(* IEC 61131-3 sources: 2026_Projet_YGO_ExcavatriceDragage/CODE/J_SUPERVISION, 7 files *)

(* ---- GVL_Troubleshooting.st ---- *)
(* ═══════════════════════════════════════════════════════════════
   🕵️‍♂️ GVL_Troubleshooting — GVL Globale de Recherche de Pannes (Orientée Fonctions & Contexte)
   ───────────────────────────────────────────────────────────────
   ⚙️ Emplacement : CODE/J_SUPERVISION/GVL_Troubleshooting.st
   🎨 Structurée par CONTEXTE GLOBAL MACHINE + FONCTIONS MÉTIER (Utilisation Opérateur).
   💬 Permet de localiser en 3 secondes l'environnement et le blocage d'une action.
   ═══════════════════════════════════════════════════════════════ *)
{attribute 'qualified_only'}
VAR_GLOBAL
    A_ContexteMachineGlobal : ST_ChainContextGlobal; // 🌐 0. Contexte Global Machine (Mode, Simu, Commande, Bypass)
    B_Inputs                : ST_HardwareImage;     // 📥 1. Image complète des entrées réelles / qualifiées / simulées
    C_Safety                : ST_SafetyChecklist;   // 🛡️ 2. Diagnostic chronologique Chaîne de Sécurité & Réarmement AU
    D_Joystick              : ST_JoystickChecklist; // 🕹️ 3. Diagnostic chronologique Bus CANopen & Homme-Mort Joystick
    E_HomingM1              : ST_HomingChecklist;   // 🎯 4. Diagnostic chronologique Homing M1 (Treuil Retenue)
    F_HomingM2              : ST_HomingChecklist;   // 🎯 5. Diagnostic chronologique Homing M2 (Treuil Benne)
    G_CycleSemiAuto         : ST_ChainCycleSemiAuto;  // 🔄 6. Séquenceur de Cycle Semi-Automatique (X0 à X13)
    H_LevageSynchroniseM1M2 : ST_ChainWinchSync;     // 🛗 7. Levage Synchronisé M1+M2 (Mode Couplé Nominal)
    I_LevageUnitaireM1      : ST_ChainWinch;         // 🛗 8. Levage Unitaire M1 (Treuil Retenue)
    J_LevageUnitaireM2      : ST_ChainWinch;         // 🛗 9. Levage Unitaire M2 (Treuil Benne)
    K_BenneOuvertureFermeture: ST_ChainBucket;        // 🪣 10. Ouverture / Fermeture Benne
    L_TranslationPontM3     : ST_ChainTranslation;   // ↔️ 11. Translation Pont M3 (Variateur AC600)
    // M_Réserve
    N_MotionM1              : ST_MotionChecklist;   // ⚙️ 13. Diagnostic chronologique Mouvement M1 (Treuil Retenue)
    O_MotionM2              : ST_MotionChecklist;   // ⚙️ 14. Diagnostic chronologique Mouvement M2 (Treuil Benne)
    P_MotionM3              : ST_MotionChecklist;   // ⚙️ 15. Diagnostic chronologique Mouvement M3 (Translation)

    // 🕵️ Trace de blocage terrain (cause priorisée + horodatage) — produite par PRG_04/05
    Q_TraceWinchM1          : ST_TraceWinch;        // 🕵️ 16. Trace blocage treuil M1 (cause priorisée + horodatage)
    R_TraceWinchM2          : ST_TraceWinch;        // 🕵️ 17. Trace blocage treuil M2 (cause priorisée + horodatage)
    S_TraceTranslation      : ST_TraceTranslation;  // ↔️ 18. Trace blocage translation M3 (cause priorisée + horodatage)
    T_Permits : ST_PermitVisibilityHMI; // Vue unique IHM/terrain des permis canoniques
END_VAR

(* ---- FB_AntiFlickerText.st ---- *)
(* ═══════════════════════════════════════════════════════════════
   🧊 FB_AntiFlickerText — Lissage anti-clignotement d'un texte IHM
   ───────────────────────────────────────────────────────────────
   📄 Doc : DOC/AF/AF_Partie-07_Interface_IHM_v2.3.md §5.3
   🎯 Responsabilité : maintient un texte warning/état un temps minimum
      avant de laisser le contenu changer, et laisse passer en direct
      (sans maintien) les messages critiques (défauts AU/puissance).
   🛡️ Sécurité : l'action de sécurité reste instantanée — ce FB ne
      retarde jamais un texte, il ne fait que stabiliser l'affichage.
      Il n'a aucun effet sur la machine.
   ═══════════════════════════════════════════════════════════════ *)
FUNCTION_BLOCK PUBLIC FB_AntiFlickerText
VAR_INPUT
    NewText      : STRING(120);  (* --> [CMD] Texte candidat à afficher *)
    ForceInstant : BOOL;         (* --> [CMD] TRUE = afficher immédiatement (défaut critique), sans maintien *)
    HoldTime     : TIME := T#500ms; (* --> [CFG] Durée de maintien min avant changement (AF-07 §5.3) *)
END_VAR
VAR_OUTPUT
    Text         : STRING(120);  (* <-- [STAT] Texte stabilisé exposé à l'IHM *)
END_VAR
VAR
    TonHold      : TON;   (* . [LOC] Temporisation de maintien *)
END_VAR

{region "§1 Lissage anti-clignotement"}
// Défaut critique : affichage immédiat, le TON est remis à zéro (aucune latence).
IF ForceInstant THEN
    Text := NewText;
    TonHold(IN := FALSE);
ELSE
    // Warning / état : le texte ne change qu'après maintien min (HoldTime).
    // Un signal qui oscille plus vite que HoldTime → texte stable.
    TonHold(IN := (NewText <> Text), PT := HoldTime);
    IF TonHold.Q THEN
        Text := NewText;
    END_IF;
END_IF;
{endregion}

(* ---- FB_CfgT330Normalizer.st ---- *)
(* ═══════════════════════════════════════════════════════════════
   🔧 FB_CfgT330Normalizer — Normalisation des réglages HAUT (T330)
   ───────────────────────────────────────────────────────────────
   🎯 Rôle : ramener DANS SON DOMAINE le couple de réglages de fin de
             course HAUT — FDC logiciel (CfgCableLimitAscent_M) et cote
             TOP homing (CfgTopSensorPos_M) — plus le plancher du
             ralentissement haut (WinchSlowdownDistanceTop_M), puis
             signaler la correction à l'IHM.
   📄 Doc : DOC/WFLOW/AUDITS/DESIGN/PLAN_T330_C3_INVARIANT_HAUT_v1.0.md (plan C3 v1.3, §2/§4)
            DOC/WFLOW/AUDITS/DESIGN/CADRAGE_T330_INVARIANT_HAUT_v1.0.md
   🛡️ Sécurité : une valeur de réglage HORS DOMAINE resterait hors domaine
             indéfiniment sans ce bloc (contre-exemple Q21 bis : FDC=9,50 m +
             TOP=12,00 m, où Δ=2,50 m ≥ 1,00 m n'active AUCUNE règle Δ).
             ⇒ R0 (clamp absolu) est INCONDITIONNELLE et EN AMONT de la règle Δ.
             Ce FB ne commande AUCUN mouvement : il corrige de la configuration.
   🧩 Dépendances : ST_WinchCfg (CfgTopSensorPos_M) · ST_CommunCfg
             (CfgCableLimitAscent_M, WinchSlowdownDistanceTop_M).
   ⚠️ Ordre d'appel : AVANT les ponts de persistance (PRG_07_Supervision §2).
             Le pont écrit la valeur CORRIGÉE dans le MÊME scan (option A / Q23)
             ⇒ aucune fenêtre NVRAM. Les mémoires internes sont amorcées depuis
             ces valeurs RESTAURÉES, jamais depuis les défauts du DUT (piège P2).
   ═══════════════════════════════════════════════════════════════ *)

FUNCTION_BLOCK FB_CfgT330Normalizer
VAR_INPUT
    // === CONTRAT STANDARD (Enable) ===
    Enable              : BOOL;  // 🟢 Autorise la normalisation (ponts de config RESTAURÉS)

    // === CONTEXTE MACHINE ===
    InHoming            : BOOL;  // 🎯 Homing en cours : cycle machine COMPLET (HX0..HX6) OU transaction de preset, M1 ou M2
END_VAR

VAR_IN_OUT
    // === RÉGLAGES HAUT À NORMALISER (référence — jamais de copie) ===
    WinchCfgM1          : ST_WinchCfg;   // 🔧 M1 = MAÎTRE du capteur haut : porte CfgTopSensorPos_M
    CommunCfg           : ST_CommunCfg;  // 🔧 Commun M1/M2 : porte CfgCableLimitAscent_M + WinchSlowdownDistanceTop_M
END_VAR

VAR_OUTPUT
    // === CONTRAT STANDARD (Ready) ===
    Ready               : BOOL;  // 🟢 Normalisation armée ce scan (Enable ET mémoires amorcées)

    // === DIAGNOSTIC / IHM ===
    Corrected           : BOOL;  // 🔧 Une correction T330 a eu lieu CE scan (impulsion d'un seul scan)
    CorrectedHeld       : BOOL;  // 🔧 Maintien du message T330 (fenêtre IHM — 1 scan serait invisible)
END_VAR

VAR CONSTANT
    // === T330 (Q1/Q2) — RÈGLES D'INGÉNIERIE, PAS DES COTES MÉTIER ===
    // NON persistantes et NON IHM (AC3) : jamais exposées, jamais RETAIN.
    CST_T330ReserveMinMargin_M : REAL := 0.40;   // Réserve minimale FDC logiciel haut / TOP homing (decision humaine, ex-1.00m)
    CST_T330SlowdownTopMin_M   : REAL := 0.50;   // Plancher du ralentissement haut (Q1)
    CST_T330FdcMin_M           : REAL := 0.00;   // Borne basse FDC (Q21)
    CST_T330FdcMax_M           : REAL := 9.60;   // Borne haute FDC (Q21/C1 : TOP<=10 et Delta>=0.4 => FDC<=9.6)
    CST_T330TopMin_M           : REAL := 1.00;   // Borne basse TOP (Q21)
    CST_T330TopMax_M           : REAL := 10.00;  // Borne haute TOP (Q21)
END_VAR

VAR
    // === T330 — MÉMOIRES NON PERSISTANTES (AC3 : ni IHM, ni RETAIN) ===
    T330PrevInit               : BOOL;  // . [LOC] Seed des mémoires effectué depuis les valeurs RESTAURÉES
    T330PrevTopSensorPos_M     : REAL;  // . [LOC] Valeur précédente TOP (détection du champ modifié par l'opérateur)
    T330PrevCableLimitAscent_M : REAL;  // . [LOC] Valeur précédente FDC (détection du champ modifié par l'opérateur)
    T330MsgHold                : TOF;   // . [LOC] Maintien du message T330 (un scan de 10 ms serait invisible à l'IHM)
END_VAR

// ═══════════════════════════════════════════════════════════════════════════════
// 🔧 T330 — COHÉRENCE DES RÉGLAGES HAUT (Q1/Q2) · plan C3 v1.3
// ───────────────────────────────────────────────────────────────────────────────
// ORDRE IMPOSÉ (Q21 bis) :  (1) R0 clamp ABSOLU inconditionnel, FDC et TOP séparément
//                        puis (2) règle Delta >= 1,00 m / slowdown >= 0,50 m.
// OPTION A (Q23) : ce bloc s'exécute AVANT les ponts de persistance, qui écrivent la
//                  valeur CORRIGÉE dans le MÊME scan (aucune fenêtre NVRAM). La
//                  référence est donc lue sur GVL_IHM.Cfg — l'état que les ponts
//                  tiennent à jour, et NON directement la NVRAM.
// AC3 : AUCUNE variable persistante ni IHM nouvelle — constantes CST_* et mémoires
//       locales uniquement. Jamais de champ de fin de course supplémentaire.
// C2/Q22 : R2 (correction du TOP) est INHIBÉE pendant le homing — sur le CYCLE COMPLET
//          (HX0..HX6), pas seulement la transaction de preset (~50 ms). Aucune mémoire
//          d'intention : au retour, si la config est toujours invalide, le REPLI NIVEAU
//          ci-dessous applique Q17 (préserver le TOP, corriger le FDC).
// ═══════════════════════════════════════════════════════════════════════════════
{region "🔧 T330 NORMALISATION"}
Corrected := FALSE;
Ready := FALSE;

// Inhibée tant que les ponts n'ont pas RESTAURÉ (sinon les défauts DUT seraient pris
// pour une saisie opérateur — piège P2 du cadrage).
IF Enable THEN

    // Seed des mémoires depuis les valeurs RESTAURÉES (jamais depuis les défauts DUT).
    IF NOT T330PrevInit THEN
        T330PrevTopSensorPos_M     := WinchCfgM1.CfgTopSensorPos_M;
        T330PrevCableLimitAscent_M := CommunCfg.CfgCableLimitAscent_M;
        T330PrevInit               := TRUE;
    END_IF;

    Ready := TRUE;

    // ─── GEL PENDANT LE HOMING (décision C2 b : « NVRAM gelée — AUCUNE écriture Cfg ») ──
    // Toutes les écritures ci-dessous (R0, R3, R1, R2) sont suspendues pendant le homing.
    // ⚠️ Ce gel couvre R1/R0/R3 AUSSI : une correction pendant un homing déplacerait la CIBLE
    // de homing (R0/R2) ou détruirait le réglage commissionné (R1) et le persisterait.
    // ⇒ À la sortie du homing, les mémoires ont suivi la saisie (bloc ci-dessous, hors gel) :
    //    il n'y a plus de FRONT, donc le REPLI NIVEAU applique R1 = Q17 (préserver le TOP). C'est
    //    exactement la décision 2c : « rien à mémoriser, on retombe dans le cas normal Q2 ».
    IF NOT InHoming THEN

    // ─── (1) R0 — CLAMP ABSOLU (Q21 bis) : non conditionné à une violation de Delta ──────
    // ⚠️ « INCONDITIONNEL » au sens de Q21 bis = non subordonné à la règle Delta. Le gel
    //    homing ci-dessus reste prioritaire (décision C2 b, motivée sécurité).
    IF CommunCfg.CfgCableLimitAscent_M < CST_T330FdcMin_M THEN
        CommunCfg.CfgCableLimitAscent_M := CST_T330FdcMin_M;
        Corrected := TRUE;
    ELSIF CommunCfg.CfgCableLimitAscent_M > CST_T330FdcMax_M THEN
        CommunCfg.CfgCableLimitAscent_M := CST_T330FdcMax_M;
        Corrected := TRUE;
    END_IF;
    IF WinchCfgM1.CfgTopSensorPos_M < CST_T330TopMin_M THEN
        WinchCfgM1.CfgTopSensorPos_M := CST_T330TopMin_M;
        Corrected := TRUE;
    ELSIF WinchCfgM1.CfgTopSensorPos_M > CST_T330TopMax_M THEN
        WinchCfgM1.CfgTopSensorPos_M := CST_T330TopMax_M;
        Corrected := TRUE;
    END_IF;

    // ─── (2) R3 — plancher du ralentissement haut ───────────────────────────────────────
    IF CommunCfg.WinchSlowdownDistanceTop_M < CST_T330SlowdownTopMin_M THEN
        CommunCfg.WinchSlowdownDistanceTop_M := CST_T330SlowdownTopMin_M;
        Corrected := TRUE;
    END_IF;

    // ─── (3) R1 / R2 — règle Delta >= 1,00 m sur les valeurs CLAMPÉES ───────────────────
    // Détection du champ MODIFIÉ : M1 (maître) et FDC commun uniquement.
    // ⛔ JAMAIS le champ M2 : il est RÉÉCRIT chaque scan par le miroir M1 (PRG_07_Supervision).
    IF (WinchCfgM1.CfgTopSensorPos_M
        - CommunCfg.CfgCableLimitAscent_M) < CST_T330ReserveMinMargin_M THEN
        IF (WinchCfgM1.CfgTopSensorPos_M <> T330PrevTopSensorPos_M)
           AND (CommunCfg.CfgCableLimitAscent_M = T330PrevCableLimitAscent_M) THEN
            // R2 — le TOP vient d'être saisi : corriger le TOP, sauf pendant le homing (C2/Q22).
            // ⚠️ Ce test est structurellement TOUJOURS VRAI ici (le gel homing englobe déjà le
            //    bloc) : il est CONSERVÉ comme marqueur nommé de la décision C2/Q22, pour qu'un
            //    déplacement futur du gel ne puisse pas réactiver R2 pendant un homing en silence.
            IF NOT InHoming THEN
                WinchCfgM1.CfgTopSensorPos_M :=
                    CommunCfg.CfgCableLimitAscent_M + CST_T330ReserveMinMargin_M;
                Corrected := TRUE;
            END_IF;
        ELSE
            // R1 (et Q17 : les deux champs ont changé, ou aucun) — PRÉSERVER le TOP,
            // corriger le FDC. C'est aussi le REPLI NIVEAU à la sortie du homing.
            CommunCfg.CfgCableLimitAscent_M :=
                WinchCfgM1.CfgTopSensorPos_M - CST_T330ReserveMinMargin_M;
            Corrected := TRUE;
        END_IF;
    END_IF;   // fin de la règle Delta (R1/R2)
    END_IF;   // ─── fin du GEL HOMING (décision C2 b) : plus aucune écriture Cfg pendant le homing

    // ─── Mémoires de front (HORS gel : suivies MÊME pendant le homing) ──────────────────
    // Indispensable : à la sortie du homing la saisie opérateur n'est plus un FRONT, donc le
    // REPLI NIVEAU ci-dessus applique R1 = Q17 (préserver le TOP, corriger le FDC). C'est la
    // décision 2c : « rien à mémoriser, on retombe dans le cas normal Q2 ».
    T330PrevTopSensorPos_M     := WinchCfgM1.CfgTopSensorPos_M;
    T330PrevCableLimitAscent_M := CommunCfg.CfgCableLimitAscent_M;

ELSE
    // Ponts non restaurés : aucune écriture Cfg, aucune mémoire amorcée.
    Ready := FALSE;
END_IF;

// Maintien IHM : une correction dure UN scan (10 ms) -> sans maintien le message serait
// invisible. TOF = conserve Q VRAI pendant PT après retombée de IN (fenêtre de maintien).
// Appelé à CHAQUE scan, y compris normalisation inhibée (la fenêtre doit pouvoir retomber).
T330MsgHold(IN := Corrected, PT := T#500ms);
CorrectedHeld := T330MsgHold.Q;
{endregion}
END_FUNCTION_BLOCK

(* ---- FB_Hmi_BannerFormatter.st ---- *)
(* ═══════════════════════════════════════════════════════════════
   🧠 FB_Hmi_BannerFormatter — Formateur du bandeau d'information IHM
   ───────────────────────────────────────────────────────────────
   📄 Doc : DOC/AF/AF_Partie-07_Interface_IHM_v2.3.md §5, §6
   🎯 Responsabilité : assemble les 4 textes du bandeau + le carrousel
      d'alarmes, expose la cause observable du blocage courant, sans
      piloter la machine.
   🛡️ Sécurité : priorité AU/puissance, SafeStop, puis interlocks métier.
      L'anti-clignotement est délégué à FB_AntiFlickerText (AF-07 §5.3).
   ═══════════════════════════════════════════════════════════════ *)
FUNCTION_BLOCK PUBLIC FB_Hmi_BannerFormatter
VAR_INPUT
    Enable               : BOOL := TRUE;   // --> [CMD] Active le formateur
    SimulationModeActive : BOOL;   // --> [TST] Mode simulation actif
    CurrentMode          : E_Mode;   // --> [CMD] Mode courant
    BothAxesCoupled      : BOOL;   // --> [HW] Treuils M1/M2 couplés
    WinchSelected        : INT; // --> [CMD] 1 = M1, 2 = M2

    // 🔄 Cycle & sous-cycles
    CycleStep            : E_AutoCycleStep;   // --> [HW] Étape cycle
    CycleStateStr        : STRING(80);   // --> [HW] Libellé détaillé de l'étape cycle (FB_CycleSemiAuto.CycleStateStr)
    CycleErrorId         : WORD;   // --> [DIAG] Code défaut cycle actif/latche (jamais 0 en AX_STAB)
    CycleStepAtError     : E_AutoCycleStep;   // --> [DIAG] Dernière étape avant le défaut (FB_CycleSemiAuto.CycleStepAtError)
    CycleChecksInhibited : BOOL;   // --> [TST] Mode essai cycle : controles procede inhibes
    MachineHomingStep        : INT;   // --> [HW] Étape guide homing machine (E_MachineHomingStep : 0..70, 60 = valide)
    MachineHomingInstruction : STRING(120);   // --> [HW] Consigne opérateur en clair produite par FB_CycleMachineHoming
    MachineHomingActionText  : STRING(120) := ''; // --> [DIAG] Consigne action operateur directe du GRAFCET homing
    MachineHomingActive      : BOOL := FALSE; // --> [HW] Cycle de homing actif (HX1..HX4)
    MachineHomingSoftLimitsOff : BOOL := FALSE; // --> [SAFE] Butees soft inhibees pendant le homing
    MachineHomingFailed      : BOOL := FALSE; // --> [DIAG] Echec ou abandon cycle homing machine
    MachineHomingLoss        : BOOL := FALSE; // --> [DIAG] Perte reference en mouvement (HomingLoss)
    MachineHomingProvisional : BOOL := FALSE; // --> [DIAG] Zero provisoire 0m HX1 actif (machine non encore calibree)
    TopHardStopLatched       : BOOL := FALSE; // --> [SAFE] Latch directionnel capteur TOP actif (montee bloquee)
    TopPositionSensorActive  : BOOL := FALSE; // --> [HW] Capteur position haute physique au contact
    WinchM1Error             : BOOL := FALSE; // --> [DIAG] Defaut commande/barriere treuil M1 (FB_Winch/Interlock)
    WinchM2Error             : BOOL := FALSE; // --> [DIAG] Defaut commande/barriere treuil M2 (FB_Winch/Interlock)
    SyncFaultLatched         : BOOL := FALSE; // --> [DIAG] Defaut synchro M1/M2 latche (Reset requis)
    BucketFaultLatched       : BOOL := FALSE; // --> [DIAG] Defaut benne latche (Reset requis)
    EncoderM1Fault           : BOOL := FALSE; // --> [DIAG] Defaut codeur M1
    EncoderM2Fault           : BOOL := FALSE; // --> [DIAG] Defaut codeur M2
    JoystickLatchedFault     : BOOL := FALSE; // --> [DIAG] Defaut joystick latche

    // 🛡️ Dérogations & particularités
    BypassGlobalActive   : BOOL;   // --> [TST] Bypass global
    CfgCorrectedT330     : BOOL;   // --> [CFG] T330 : correction automatique d'un reglage haut (fenetre de maintien)
    BypassWinchM1Active  : BOOL;   // --> [TST] Bypass treuil M1
    BypassWinchM2Active  : BOOL;   // --> [TST] Bypass treuil M2
    BypassTranslation    : BOOL;   // --> [TST] Bypass translation
    BypassSyncActive     : BOOL;   // --> [TST] Bypass synchro
    SyncDegradedActive   : BOOL;   // --> [TST] Synchro bridée
    LegalLimitReached    : BOOL;   // --> [SAFE] Limite légale atteinte
    ModeChangePendingBlocked : BOOL;   // --> [DIAG] Bascule de mode refusée (treuils non à l'arrêt)
    ModeChangeBlockReason    : STRING(40); // --> [DIAG] Motif du blocage de bascule (ex. "Chgt mode refuse : contacteur M1")

    // 🎮 Sécurité, causes et intention de direction
    EmergencyChainClosed : BOOL;   // --> [SAFE] Chaîne AU fermée
    PowerContactorEngaged: BOOL;   // --> [SAFE] Contacteur puissance
    PowerCutOffActiveAny : BOOL;   // --> [SAFE] Coupure puissance active
    SafeStopActive       : BOOL; // --> [SAFE] Agrégat M1/M2 par OR — tout SafeStop affiché (bandeau conservateur)
    DescendPermit        : BOOL; // --> [SAFE] Agrégat M1/M2 par AND
    AscentPermit         : BOOL; // --> [SAFE] Agrégat M1/M2 par AND
    BucketIsOpen         : BOOL;   // --> [HW] Benne ouverte
    BucketIsClosed       : BOOL;   // --> [HW] Benne fermee (montee non bridée)
    DiveActive           : BOOL;   // --> [HW] Plongée active
    TopLimitReached      : BOOL; // --> [SAFE] Agrégat M1/M2 par OR — toute limite haute affichée
    WinchBothMotionDirection : INT;   // --> [CMD] Direction demandée couplée
    M1LogicRequestDirection     : INT;   // --> [CMD] Direction logique M1
    M2LogicRequestDirection     : INT;   // --> [CMD] Direction logique M2
    CycleRequestDirection      : INT;   // --> [CMD] Direction cycle
    DeadmanArmed         : BOOL;   // --> [SAFE] Homme-mort armé
    JoystickAtNeutral    : BOOL;   // --> [HW] Joystick au neutre
    ArmingPermitDenied   : BOOL;   // --> [DIAG] Appui homme-mort refusé (ArmingPermit=FALSE)
    ArmingBlockedReason  : E_ArmingBlockReason; // --> [DIAG] Motif précis du refus d'armement
    CycleAutoBusy        : BOOL;   // --> [HW] Cycle auto actif
    CycleElapsed_Min     : INT;   // --> [DIAG] Minutes ecoulees du cycle EN COURS (FB_CycleSemiAuto.CurrentCycleElapsed_Min) — affichees seulement si CycleAutoBusy
    CycleElapsed_S       : INT;   // --> [DIAG] Secondes ecoulees du cycle EN COURS, 0..59 (FB_CycleSemiAuto.CurrentCycleElapsed_S)
    M3AtP1               : BOOL;   // --> [STAT] M3 positionné stable au Point 1 (conservé, compat)
    M3StatusText         : STRING(80);   // --> [STAT] T249-B : texte statut position M3 (PRG_05) — "M3 a P1", "M3 entre P2 et P1 -> Maintenance"...
    TranslationMotionErrorId       : WORD;   // --> [DIAG] Code défaut MOUVEMENT M3 (FB_Translation.Fault.ErrorId) : bit0 frein, bit3 variateur AC600, bit6 limite extrême
    TranslationFinalInterlockErrorId : WORD; // --> [DIAG] Code défaut barrière finale M3 (frein / redémarrage)
    WinchDescentLockedByM3 : BOOL;   // --> [STAT] T249-A : descente M1/M2 verrouillée, chariot M3 pas à P1/Maintenance (info, pas alarme)
    M3AtTremieStable     : BOOL;   // --> [STAT] M3 arrêté stable à la Trémie (latch FdC) — mode benne dispo, prioritaire sur WinchDescentLockedByM3

    // 🚨 Bandeau d'alarme défilant (§5) — diagnostics safety et ErrorId machine entière
    WinchM1Safety        : ST_SafetyWinch;       // --> [SAFE] Diagnostic sécurité treuil M1
    WinchM2Safety        : ST_SafetyWinch;       // --> [SAFE] Diagnostic sécurité treuil M2
    TranslationSafety    : ST_SafetyTranslation; // --> [SAFE] Diagnostic sécurité translation M3
    BucketErrorId        : WORD;   // --> [DIAG] Code défaut benne (FB_Bucket.ErrorId)
    SyncErrorId          : WORD;   // --> [DIAG] Code défaut synchro M1/M2 (FB_WinchSync.ErrorId)
    SyncContactorDiag    : ST_SyncContactorDiag;   // --> [DIAG] Discordance contacteurs M1/M2 décodée (FB_SyncContactor PRG_06 §2quinquies)
    DiveErrorId          : WORD;   // --> [DIAG] Code défaut plongée (FB_DiveSearch.ErrorId)
    ExtractionErrorId    : WORD;   // --> [DIAG] Code défaut extraction (FB_ExtractionAssist.ErrorId)
    EmergencyErrorId     : WORD;   // --> [DIAG] Code défaut chaîne AU (FB_Safety_EmergencyManagement.Diag.ErrorId)
    RedundancyTestFailed : BOOL;   // --> [DIAG] Defaut redondance contacteurs AU (lisee -> message explicite)
    EmergencyArmingFailed: BOOL;   // --> [DIAG] Echec rearmement contacteur AU (lisee -> message explicite)
    ArmingSeqStep        : INT;    // --> [DIAG] Etape sequence rearmement AU (0=IDLE..6=Confirm) — front descendant = abandon
    LastAbortCause       : WORD;   // --> [DIAG] Cause du dernier abandon de sequence AU (message explicite cause+action)
    Reset                : BOOL;   // --> [CMD] Front acquittement defauts (FaultMachineReset_IHM) — efface le message d'abandon verrouillé
    AlarmHoldTime        : TIME := T#1s; // --> [CFG] Durée d'affichage par message du carrousel
    Network              : ST_NetworkDiagHMI; // --> [DIAG] Diagnostic réseau, bus et modules E/S
END_VAR
VAR_OUTPUT
    Banner               : ST_HmiBanner;   // <-- [STAT] Bandeau IHM assemblé
END_VAR
VAR
    PrefixContext        : STRING(20);   // . [LOC] Préfixe RÉEL/SIMU
    ModeStr              : STRING(30);   // . [LOC] Libellé mode
    CouplingStr          : STRING(30);   // . [LOC] Libellé couplage
    ElapsedSuffixStr     : STRING(20);  // . [LOC] Suffixe chrono du cycle en cours, format ' MMminSSs' (deux chiffres par champ)
    CurrentDirection     : INT;   // . [LOC] Direction courante
    DirectionBlocked     : BOOL; // . [LOC] Interlock métier : mouvement demandé mais permit absent
    AnyBypassActive      : BOOL;   // . [LOC] Au moins un bypass actif
    PowerOrChainFault    : BOOL; // . [LOC] Défaut chaîne AU ou contacteur puissance absent
    HardwareModuleOrBusFault : BOOL; // . [LOC] Défaut matériel module E/S ou bus actif
    CriticalActionActive : BOOL; // . [LOC] Défaut/interlock critique : affiché immédiatement (sans maintien)
    SpecialConditionCandidate : STRING(120);   // . [LOC] Texte condition spéciale
    OperatorActionCandidate   : STRING(120);   // . [LOC] Texte action opérateur
    StepAtErrorStr            : STRING(40);   // . [LOC] Libellé de l'étape d'origine du défaut
    CycleFaultCauseStr        : STRING(120);  // . [LOC] Cause cycle décodée pour acquittement terrain
    WinchRootCauseStr         : STRING(32);   // . [LOC] Cause racine winch affichée en repli AX_STAB
    WinchRootTagStr           : STRING(4);    // . [LOC] Étiquette treuil concerné (M1/M2) de la cause racine
    WinchRootCauseLbl         : STRING(20);   // . [LOC] Libellé court de la cause racine winch
    WinchRootMaskId           : WORD;         // . [LOC] Masque latché du treuil retenu (M1 prioritaire, sinon M2)
    CycleFaultActive          : BOOL;         // . [LOC] Repli AX_STAB sur défaut cycle (cause latchee presente)
    CycleFaultMsgStr          : STRING(120);  // . [LOC] Message [CYCLE] de repli : cause cycle + cause racine
    AntiFlickSpecial     : FB_AntiFlickerText; // * [INST] §3 Condition spéciale (warning → maintenu)
    AntiFlickOperator    : FB_AntiFlickerText; // * [INST] §4 Action opérateur (critique → direct, warning → maintenu)
    LastAbortEdge        : F_TRIG; // . [LOC] Front descendant ArmingSeqStep (abandon de sequence AU)
    ArmingInProgress     : BOOL; // . [LOC] Sequence AU en cours (ArmingSeqStep <> 0)
    ResetEdge            : R_TRIG; // . [LOC] Front montant Reset (acquittement defauts)
    ArmStartEdge         : R_TRIG; // . [LOC] Front montant ArmingInProgress (nouvelle sequence AU)
    TonAbortHold         : TON; // . [LOC] Maintien du message d'abandon AU (causes non latched)
    AbortMsgActive       : BOOL; // . [LOC] Message d'abandon AU affiché (fenêtre de maintien)
    AbortMsgLatched      : BOOL; // . [LOC] Message d'abandon verrouillé jusqu'à Reset (causes sans latch)
    AbortMsgText         : STRING(120); // . [LOC] Texte cause+action du dernier abandon AU
    SeqReachedConfirm    : BOOL; // . [LOC] La sequence AU a atteint l'etape 6 (confirmation) -> distingue SUCCES d'un ABANDON
    TonAlarmBanner       : TON; // . [LOC] §5 Tempo de maintien par message du carrousel
    AlarmArray           : ARRAY[0..49] OF STRING(120); // . [LOC] §5 Messages actifs collectés ce scan
    AlarmCount           : INT; // . [LOC] §5 Nombre de messages actifs
    BannerSyncContactorWhich : STRING(80); // . [LOC] §5 Libellé du contacteur M1/M2 en discordance
    AlarmIndex           : INT; // . [LOC] §5 Index courant du carrousel (0-based)
    i                    : INT; // . [LOC] Index de boucle
    TonBootInhibit       : TON; // . [LOC] Garde au démarrage (inhibition fausses alarmes réseau 4s)
    TofFaultLocalIo      : TOF; // . [LOC] Anti-bagotement Local_Digital_IO (1.5s)
    TofFaultVh0800       : TOF; // . [LOC] Anti-bagotement VH_0800END (1.5s)
    TofFaultVh0808       : TOF; // . [LOC] Anti-bagotement VH_0808ETP (1.5s)
    TofFaultVh0008Er     : TOF; // . [LOC] Anti-bagotement VH_0008ER (1.5s)
    TofFaultVh0008Er1    : TOF; // . [LOC] Anti-bagotement VH_0008ER_1 (1.5s)
    TofFaultCanBus       : TOF; // . [LOC] Anti-bagotement bus CANopen (1.5s)
    TofFaultJoy1         : TOF; // . [LOC] Anti-bagotement Joystick JOY1 (1.5s)
    TofFaultEcatBus      : TOF; // . [LOC] Anti-bagotement bus EtherCAT (1.5s)
    TofFaultEncM1        : TOF; // . [LOC] Anti-bagotement EtherCAT Encoder M1 (1.5s)
    TofFaultEncM2        : TOF; // . [LOC] Anti-bagotement EtherCAT Encoder M2 (1.5s)
    TofFaultVarM3        : TOF; // . [LOC] Anti-bagotement EtherCAT Variateur M3 (1.5s)
    LocalIoValid         : BOOL; // . [LOC] Validité filtrée Local_Digital_IO (DI8/DO8)
    Vh0800Valid          : BOOL; // . [LOC] Validité filtrée VH_0800END (DI8)
    Vh0808Valid          : BOOL; // . [LOC] Validité filtrée VH_0808ETP (DI8/DO8)
    Vh0008ErValid        : BOOL; // . [LOC] Validité filtrée VH_0008ER (DO8 Relais Freins/Kobold)
    Vh0008Er1Valid       : BOOL; // . [LOC] Validité filtrée VH_0008ER_1 (DO8 Relais AU/PowerKeepAlive)
    CanBusValid          : BOOL; // . [LOC] Validité filtrée Bus CANopen
    Joy1Valid            : BOOL; // . [LOC] Validité filtrée Joystick JOY1
    EcatBusValid         : BOOL; // . [LOC] Validité filtrée Bus EtherCAT
    EncM1Valid           : BOOL; // . [LOC] Validité filtrée Encoder M1
    EncM2Valid           : BOOL; // . [LOC] Validité filtrée Encoder M2
    VarM3Valid           : BOOL; // . [LOC] Validité filtrée Variateur M3
    HistoM1              : WORD; // . [LOC] §5 [HISTO] M1 : LatchedId AND NOT ErrorId (défauts latched passés)
    HistoM2              : WORD; // . [LOC] §5 [HISTO] M2 : LatchedId AND NOT ErrorId (défauts latched passés)
    HistoM3              : WORD; // . [LOC] §5 [HISTO] M3 : LatchedId AND NOT ErrorId (défauts latched passés)
    RearmEdge            : R_TRIG; // . [LOC] Front du réarmement puissance (contacteur)
    TonRearmWindow       : TON;    // . [LOC] Fenêtre transitoire post-réarmement (durée bornée)
    RearmWindowActive    : BOOL;   // . [LOC] Fenêtre post-réarmement en cours
    NetworkSurveillanceActive : BOOL; // . [LOC] Surveillance réseau/ES armée (hors fenêtre transitoire attendue)
END_VAR
VAR CONSTANT
    CST_BannerHoldTime   : TIME := T#500ms; // . [LOC] Anti-clignotement warnings/états (AF-07 §5.3)
    CST_AbortHoldTime    : TIME := T#5s; // . [LOC] Maintien message d'abandon AU
    CST_NbMaxAlarmes     : INT := 50; // . [LOC] Taille du carrousel d'alarmes (AF-07 §6)
    // ⏱️ Durée de la fenêtre transitoire post-réarmement, alignée sur la garde de démarrage :
    // pendant ce délai les esclaves peuvent légitimement ne pas être encore opérationnels.
    // C'est une BORNE : passé ce délai, un défaut réseau réel est de nouveau affiché.
    CST_RearmInhibitTime : TIME := T#4s; // . [LOC] Fenêtre transitoire post-réarmement puissance
    // 🔑 Bit 6 de ST_SafetyWinch.ErrorId = cause « Limite basse cable atteinte » (vue LIVE,
    // Latching := FALSE, FB_Safety_Winch.st:318-325). Le DUT ST_SafetyWinch n'expose aucun
    // champ nommé pour cette cause : le bit est nommé ici plutôt qu'écrit en clair.
    // ⚠️ Ne JAMAIS lire WinchMxSafety.CableLimitDescent à la place : ce champ est une
    // comparaison BRUTE de position, sans bypass ni mode référencement
    // (FB_WinchStateProjection.st:217-218/230/257) — il resterait vrai sous
    // BypassCableLimitSwitch (MAINT_N2) alors que la cause safety est levée.
    CST_WinchErrorIdCableLimitDescent : WORD := 16#0040; // . [LOC] Bit 6 ErrorId : limite basse cable
END_VAR

IF NOT Enable THEN
    Banner.GlobalContextText     := '';
    Banner.SequenceProgressText  := '';
    Banner.SpecialConditionText  := '';
    Banner.OperatorActionText    := '';
    Banner.PositionM3Text        := '';
    Banner.AlarmBanner.HasAlarm  := FALSE;
    Banner.AlarmBanner.Text      := '';
    Banner.AlarmBanner.Index     := 0;
    Banner.AlarmBanner.Count     := 0;
    FOR i := 0 TO 49 DO
        Banner.AlarmBanner.AlarmArray[i] := '';
    END_FOR;
    TonAlarmBanner(IN := FALSE);
    TonBootInhibit(IN := FALSE);
    TonRearmWindow(IN := FALSE);
    RearmEdge(CLK := FALSE);
    RearmWindowActive := FALSE;
    NetworkSurveillanceActive := FALSE;
    TofFaultLocalIo(IN := FALSE);
    TofFaultVh0800(IN := FALSE);
    TofFaultVh0808(IN := FALSE);
    TofFaultVh0008Er(IN := FALSE);
    TofFaultVh0008Er1(IN := FALSE);
    TofFaultCanBus(IN := FALSE);
    TofFaultJoy1(IN := FALSE);
    TofFaultEcatBus(IN := FALSE);
    TofFaultEncM1(IN := FALSE);
    TofFaultEncM2(IN := FALSE);
    TofFaultVarM3(IN := FALSE);
    RETURN;
END_IF;

// ⏱️ Garde au démarrage (inhibition 4s pendant init des bus et équipements)
TonBootInhibit(IN := Enable, PT := T#4s);

// ⏱️ Fenêtre transitoire de réarmement puissance : à chaque front du contacteur, les esclaves
// peuvent légitimement publier une perte de liaison pendant quelques secondes. La fenêtre est
// BORNÉE (CST_RearmInhibitTime) : hors de celle-ci, un défaut réseau réel reste affiché.
RearmEdge(CLK := PowerContactorEngaged);
IF RearmEdge.Q THEN
    RearmWindowActive := TRUE;
END_IF;
TonRearmWindow(IN := RearmWindowActive, PT := CST_RearmInhibitTime);
IF TonRearmWindow.Q THEN
    RearmWindowActive := FALSE;
END_IF;

// 🛡️ Surveillance réseau armée hors des phases où l'absence de bus est ATTENDUE :
// démarrage CPU (garde ci-dessus) et réarmement puissance (fenêtre ci-dessus).
// Rien d'autre n'est masqué : la chaîne AU, les sécurités et les défauts métier ne passent pas ici.
NetworkSurveillanceActive := TonBootInhibit.Q AND NOT RearmWindowActive;

// 🌊 Filtrage anti-bagotement (TOF 1.5s sur perte de validité)
TofFaultLocalIo(IN := (NOT Network.InputModules.LocalDigitalIoOk) AND NetworkSurveillanceActive, PT := T#1.5s);
TofFaultVh0800(IN := (NOT Network.InputModules.Vh0800EndOk) AND NetworkSurveillanceActive, PT := T#1.5s);
TofFaultVh0808(IN := (NOT Network.InputModules.Vh0808EtpOk) AND NetworkSurveillanceActive, PT := T#1.5s);
TofFaultVh0008Er(IN := (NOT Network.InputModules.Vh0008ErOk) AND NetworkSurveillanceActive, PT := T#1.5s);
TofFaultVh0008Er1(IN := (NOT Network.InputModules.Vh0008Er1Ok) AND NetworkSurveillanceActive, PT := T#1.5s);
TofFaultCanBus(IN := (NOT Network.BusCanOpen.Operational) AND NetworkSurveillanceActive, PT := T#1.5s);
TofFaultJoy1(IN := (NOT Network.Joystick.Operational) AND NetworkSurveillanceActive, PT := T#1.5s);
TofFaultEcatBus(IN := (NOT Network.BusEthercat.Operational) AND NetworkSurveillanceActive, PT := T#1.5s);
TofFaultEncM1(IN := (NOT Network.EncoderM1.Operational) AND NetworkSurveillanceActive, PT := T#1.5s);
TofFaultEncM2(IN := (NOT Network.EncoderM2.Operational) AND NetworkSurveillanceActive, PT := T#1.5s);
TofFaultVarM3(IN := (NOT Network.VariateurM3.Operational) AND NetworkSurveillanceActive, PT := T#1.5s);

LocalIoValid   := NOT TofFaultLocalIo.Q;
Vh0800Valid    := NOT TofFaultVh0800.Q;
Vh0808Valid    := NOT TofFaultVh0808.Q;
Vh0008ErValid  := NOT TofFaultVh0008Er.Q;
Vh0008Er1Valid := NOT TofFaultVh0008Er1.Q;
CanBusValid    := NOT TofFaultCanBus.Q;
Joy1Valid      := NOT TofFaultJoy1.Q;
EcatBusValid   := NOT TofFaultEcatBus.Q;
EncM1Valid     := NOT TofFaultEncM1.Q;
EncM2Valid     := NOT TofFaultEncM2.Q;
VarM3Valid     := NOT TofFaultVarM3.Q;

{region "§1 Contexte global"}
// ═══════════════════════════════════════════════════════════════
// 1. CONTEXTE GLOBAL — aucun numéro d'étape ici
// Format (AF-07 §5.1) : [RÉEL/SIMU] [MODE] [COUPLAGE]
// ═══════════════════════════════════════════════════════════════
IF SimulationModeActive THEN
    PrefixContext := '[SIMULATION] ';
ELSE
    PrefixContext := '[RÉEL] ';
END_IF;

CASE CurrentMode OF
    E_Mode.DISABLE:  ModeStr := '[DÉSACTIVÉ]';
    E_Mode.MAINT_N1: ModeStr := '[MAINT_N1]';
    E_Mode.MAINT_N2: ModeStr := '[MAINT_N2]';
    E_Mode.SEMI_AUTO: ModeStr := '[SEMI-AUTO]';
ELSE
    ModeStr := '[MODE INCONNU]';
END_CASE;

IF CurrentMode = E_Mode.SEMI_AUTO THEN
    CouplingStr := ' [CYCLE AUTO]';
ELSIF BothAxesCoupled THEN
    CouplingStr := ' [M1+M2 COUPLÉS]';
ELSIF WinchSelected = 1 THEN
    CouplingStr := ' [M1 SEUL]';
ELSIF WinchSelected = 2 THEN
    CouplingStr := ' [M2 SEUL]';
ELSE
    CouplingStr := ' [AUCUN AXE]';
END_IF;
// Assemblage par ACCUMULATION sur le champ cible (STRING(120)) plutot que par CONCAT imbrique :
// le resultat est identique en CODESYS (c'est la taille du champ cible qui gouverne), mais il ne
// depend plus de la taille declaree des fragments intermediaires. Un CONCAT imbrique de fragments
// STRING(20)/STRING(30)/STRING(30) est plafonne a 30 caracteres par le compilateur de test, qui
// fait rendre a CONCAT le maximum de la taille de ses arguments : le mode affiche ressortait
// ampute ('[SIMULATION] [SEMI-AUTO] [CYCL', 'CYCLE AUTO]' perdu) sur le harnais CI.
Banner.GlobalContextText := PrefixContext;
Banner.GlobalContextText := CONCAT(Banner.GlobalContextText, ModeStr);
Banner.GlobalContextText := CONCAT(Banner.GlobalContextText, CouplingStr);

// ⏱️ Chronomètre du cycle EN COURS, accolé au bandeau mode (format MMminSSs, ex. '09min05s').
// • Producteur unique de la valeur : FB_CycleSemiAuto (CurrentCycleElapsed_Min/_S) ; le formateur
//   ne recalcule RIEN et ne lit aucun global : les deux entiers arrivent par VAR_INPUT
//   (cablés par PRG_07_Supervision.st sur GVL_IHM.CycleSemiAuto.State).
// • Portillon : CycleAutoBusy = Lifecycle.Busy du séquenceur (PRG_07:758). Hors cycle il est FALSE
//   (PRG_03_Modes_Cycle.st:471 et :544 hors SEMI_AUTO, FB_CycleSemiAuto.st:1585 en AX18 et :1621 en
//   AX_STAB) et le chrono est remis à zéro (PRG_03_Modes_Cycle.st:490-494 / :565-569) : aucune durée
//   figée d'un cycle précédent ne peut donc s'afficher à l'arrêt.
// • Pire cas borné : 37 car. de base + 1 espace + 3 chiffres de minutes (CycleRunTimer armé PT=T#12h
//   -> 720 min maximum) + 'min' + 2 chiffres de secondes + 's' = 47 car., contre STRING(120) pour
//   GlobalContextText (ST_HmiBanner.st:10). Même si les minutes n'étaient pas bornées par le TON
//   (INT complet, 11 car.), le total resterait à 55 car. : aucune troncature possible.
IF CycleAutoBusy THEN
    IF CycleElapsed_Min < 10 THEN
        ElapsedSuffixStr := CONCAT(' 0', CONCAT(INT_TO_STRING(CycleElapsed_Min), 'min'));
    ELSE
        ElapsedSuffixStr := CONCAT(' ', CONCAT(INT_TO_STRING(CycleElapsed_Min), 'min'));
    END_IF;
    IF CycleElapsed_S < 10 THEN
        ElapsedSuffixStr := CONCAT(ElapsedSuffixStr, CONCAT('0', CONCAT(INT_TO_STRING(CycleElapsed_S), 's')));
    ELSE
        ElapsedSuffixStr := CONCAT(ElapsedSuffixStr, CONCAT(INT_TO_STRING(CycleElapsed_S), 's'));
    END_IF;
    Banner.GlobalContextText := CONCAT(Banner.GlobalContextText, ElapsedSuffixStr);
END_IF;
{endregion}

{region "§1bis Repli defaut (etape origine)"}
// ═══════════════════════════════════════════════════════════════
// 🧊 REPLI DÉFAUT (AX_STAB) — étape d'ORIGINE du défaut.
// Calculé AVANT §2 et §4 car deux champs du bandeau l'utilisent :
//   - §2 Progression : « Cycle: STABILISATION (defaut a AX7) » — en repli on n'est PLUS
//     a AX7 : le champ doit situer l'origine SANS laisser croire qu'on y est encore ;
//   - §4 Action opérateur : « [CYCLE]AX7:cause(cause racine)>Repr/Abandon ».
// ═══════════════════════════════════════════════════════════════
CycleFaultActive := (CycleStep = E_AutoCycleStep.AX_STAB) AND (CycleErrorId <> 0);
StepAtErrorStr   := '';
IF CycleFaultActive THEN
    CASE CycleStepAtError OF
        E_AutoCycleStep.AX0_REPOS: StepAtErrorStr := 'X0';
        E_AutoCycleStep.AX1_INIT: StepAtErrorStr := 'X1';
        E_AutoCycleStep.AX2_TRANSLATE_P1: StepAtErrorStr := 'X2';
        E_AutoCycleStep.AX3_OPEN_BUCKET: StepAtErrorStr := 'X3';
        E_AutoCycleStep.AX4_DESCEND_DIVING: StepAtErrorStr := 'AX4';
        E_AutoCycleStep.AX5_KOBOLD_INIT: StepAtErrorStr := 'AX5';
        E_AutoCycleStep.AX6_SEARCH_IMMERSION: StepAtErrorStr := 'AX6';
        E_AutoCycleStep.AX7_SEARCH_BOTTOM: StepAtErrorStr := 'AX7';
        E_AutoCycleStep.AX8_BOTTOM_CONFIRMED: StepAtErrorStr := 'AX8';
        E_AutoCycleStep.AX_DIVING_RETRY: StepAtErrorStr := 'RETRY';
        E_AutoCycleStep.AX9_RAISE_OFF_BOTTOM: StepAtErrorStr := 'AX9';
        E_AutoCycleStep.AX10_CLOSE_BUCKET: StepAtErrorStr := 'AX10';
        E_AutoCycleStep.AX10B_RACCORDEMENT_P1: StepAtErrorStr := 'AX10b';
        E_AutoCycleStep.AX11_CTRL_ASCENT: StepAtErrorStr := 'AX11';
        E_AutoCycleStep.AX12_LOADED_ASCENT: StepAtErrorStr := 'AX12';
        E_AutoCycleStep.AX13_DRAIN_PAUSE: StepAtErrorStr := 'AX13';
        E_AutoCycleStep.AX14_TRANSLATE_DUMP: StepAtErrorStr := 'AX14';
        E_AutoCycleStep.AX15A_DUMP_ARRIVE: StepAtErrorStr := 'AX15a';
        E_AutoCycleStep.AX15B_DUMP_OPEN: StepAtErrorStr := 'AX15b';
        E_AutoCycleStep.AX15C_DUMP_REPOSITION: StepAtErrorStr := 'AX15c';
        E_AutoCycleStep.AX18_DONE_SYNC: StepAtErrorStr := 'AX18';
        E_AutoCycleStep.AX_STAB: StepAtErrorStr := 'STAB';
        ELSE
            StepAtErrorStr := '?';
    END_CASE;
END_IF;
{endregion}

{region "§2 Progression"}
// ═══════════════════════════════════════════════════════════════
// 2. PROGRESSION — le numéro et l'étape restent exclusivement ici
// Format (AF-07 §5.1) : Macro: <Cycle> > Sous-cycle: <Étape>
// ═══════════════════════════════════════════════════════════════
// Guide homing machine : source unique = FB_CycleMachineHoming (1 texte par étape).
// Prioritaire tant que non valide (SEMI_AUTO est de toute façon interdit sans MachineHomed).
IF (MachineHomingStep > 0) AND (MachineHomingStep <> 60) THEN
    Banner.SequenceProgressText := CONCAT('Homing: ', MachineHomingInstruction);
ELSIF CurrentMode = E_Mode.SEMI_AUTO THEN
    // Repli defaut : on n'est PLUS a l'etape d'origine — on est en STABILISATION. Le champ
    // situe l'origine du defaut sans laisser croire qu'on y est encore.
    IF CycleFaultActive THEN
        Banner.SequenceProgressText := CONCAT('Cycle: STABILISATION (defaut a ',
                                     CONCAT(StepAtErrorStr, ')'));
    // Sinon : détail de l'étape (FB_CycleSemiAuto.CycleStateStr) prioritaire ; label court en fallback.
    ELSIF CycleStateStr <> '' THEN
        Banner.SequenceProgressText := CONCAT('Cycle: ', CycleStateStr);
    ELSE
        CASE CycleStep OF
            E_AutoCycleStep.AX0_REPOS: Banner.SequenceProgressText := 'Cycle: PRÉPARATION';
            E_AutoCycleStep.AX1_INIT: Banner.SequenceProgressText := 'Cycle: CONDITIONS INITIALES';
            E_AutoCycleStep.AX2_TRANSLATE_P1: Banner.SequenceProgressText := 'Cycle: TRANSLATION P1';
            E_AutoCycleStep.AX3_OPEN_BUCKET: Banner.SequenceProgressText := 'Cycle: OUVERTURE BENNE';
            E_AutoCycleStep.AX4_DESCEND_DIVING: Banner.SequenceProgressText := 'Cycle: PLONGÉE PALIER 4';
            E_AutoCycleStep.AX5_KOBOLD_INIT: Banner.SequenceProgressText := 'Cycle: INIT KOBOLD';
            E_AutoCycleStep.AX6_SEARCH_IMMERSION: Banner.SequenceProgressText := 'Cycle: RECHERCHE IMMERSION';
            E_AutoCycleStep.AX7_SEARCH_BOTTOM: Banner.SequenceProgressText := 'Cycle: RECHERCHE FOND';
            E_AutoCycleStep.AX8_BOTTOM_CONFIRMED: Banner.SequenceProgressText := 'Cycle: FOND CONFIRMÉ';
            E_AutoCycleStep.AX_DIVING_RETRY: Banner.SequenceProgressText := 'Cycle: REPRISE PLONGÉE';
            E_AutoCycleStep.AX9_RAISE_OFF_BOTTOM: Banner.SequenceProgressText := 'Cycle: MONTEE SYNCHRONISEE - RETENDRE CABLES';
            E_AutoCycleStep.AX10_CLOSE_BUCKET: Banner.SequenceProgressText := 'Cycle: FERMETURE BENNE';
            E_AutoCycleStep.AX10B_RACCORDEMENT_P1: Banner.SequenceProgressText := 'Cycle: RACCORDEMENT P1 AVANT MONTEE';
            E_AutoCycleStep.AX11_CTRL_ASCENT: Banner.SequenceProgressText := 'Cycle: MONTÉE CONTRÔLE';
            E_AutoCycleStep.AX12_LOADED_ASCENT: Banner.SequenceProgressText := 'Cycle: REMONTÉE CHARGÉE';
            E_AutoCycleStep.AX13_DRAIN_PAUSE: Banner.SequenceProgressText := 'Cycle: ÉGOUTTAGE';
            E_AutoCycleStep.AX14_TRANSLATE_DUMP: Banner.SequenceProgressText := 'Cycle: TRANSLATION TRÉMIE';
            E_AutoCycleStep.AX15A_DUMP_ARRIVE, E_AutoCycleStep.AX15B_DUMP_OPEN: Banner.SequenceProgressText := 'Cycle: VIDAGE BENNE';
            E_AutoCycleStep.AX15C_DUMP_REPOSITION: Banner.SequenceProgressText := 'Cycle: VIDAGE BENNE';
            E_AutoCycleStep.AX18_DONE_SYNC: Banner.SequenceProgressText := 'Cycle: TERMINÉ - ALLER P1';
            E_AutoCycleStep.AX_STAB: Banner.SequenceProgressText := 'Cycle: STABILISATION';
        ELSE
            Banner.SequenceProgressText := 'Cycle: ÉTAPE EN COURS';
        END_CASE;
    END_IF;
ELSIF CurrentMode = E_Mode.MAINT_N1 OR CurrentMode = E_Mode.MAINT_N2 THEN
    Banner.SequenceProgressText := 'Manuel: PILOTAGE DIRECT';
ELSE
    Banner.SequenceProgressText := 'Machine: ARRÊTÉE';
END_IF;
{endregion}

{region "§2bis Position M3"}
// État indépendant : ne participe pas aux arbitrages des quatre champs historiques
// ni au carrousel des défauts. Texte statut position M3 calculé par PRG_05 (T249-B) :
// jeton "at position" sur front capteur, sinon zone entre 2 capteurs (SensorsWord),
// + suffixe sens de déplacement. Niveau INFO, jamais alarme.
Banner.PositionM3Text := M3StatusText;
{endregion}

{region "§3 Condition spéciale"}
// ═══════════════════════════════════════════════════════════════
// 3. CONDITION SPÉCIALE — un seul indicateur bypass/dérogation
// Format (AF-07 §5.1) : ATTENTION: <Dérogation / Bridage / Alerte>
// 🧊 Warning → maintenu min (anti-clignotement), jamais critique.
// ⚠️ La simulation n'est PAS un bypass : elle n'apparaît que dans le
//    contexte global (champ 1), jamais ici.
// ═══════════════════════════════════════════════════════════════
AnyBypassActive := BypassGlobalActive
                OR BypassWinchM1Active
                OR BypassWinchM2Active
                OR BypassTranslation
                OR BypassSyncActive;
IF ModeChangePendingBlocked AND ModeChangeBlockReason <> '' THEN
    // Bascule de mode refusée : motif prioritaire (info opérateur, ex. "Chgt mode refuse : contacteur M1").
    SpecialConditionCandidate := ModeChangeBlockReason;
ELSIF CycleChecksInhibited THEN
    SpecialConditionCandidate := 'ESSAI CYCLE : CONTROLES INHIBES';
ELSIF TopHardStopLatched THEN
    SpecialConditionCandidate := 'ATTENTION: Capteur TOP franchi - redescendre';
ELSIF MachineHomingProvisional THEN
    SpecialConditionCandidate := 'ATTENTION: Ref 0m PROVISOIRE - Non calibre';
ELSIF AnyBypassActive THEN
    SpecialConditionCandidate := 'ATTENTION: Bypass actif';
ELSIF SyncDegradedActive THEN
    SpecialConditionCandidate := 'ATTENTION: Synchro bridée';
ELSIF LegalLimitReached THEN
    SpecialConditionCandidate := 'ATTENTION: Limite légale';
ELSIF M3AtTremieStable THEN
    // A la Tremie, le mode benne (WinchSel=2) reste dispo (exempte du verrou T249-A,
    // commit bb2bf240) -> priorite sur le message descente verrouillee ci-dessous, qui
    // etait le seul affiche a la Tremie et faisait croire a l'operateur que TOUT etait
    // bloque, y compris la benne (REX MES 2026-09-04).
    SpecialConditionCandidate := 'M3 a la Tremie : mode benne actif (ouverture/fermeture disponible)';
ELSIF WinchDescentLockedByM3 THEN
    // T249-A : verrou GENERAL en MAINT (pas seulement DumpAtTremie) — sans ce message
    // l'operateur ne comprend pas pourquoi la descente est refusee (REX MES 2026-09-04).
    SpecialConditionCandidate := 'Descente treuil verrouillee : chariot M3 pas a P1/Maintenance';
ELSE
    SpecialConditionCandidate := '';
END_IF;

AntiFlickSpecial(NewText := SpecialConditionCandidate, ForceInstant := FALSE, HoldTime := CST_BannerHoldTime);
Banner.SpecialConditionText := AntiFlickSpecial.Text;
{endregion}

{region "§4 Action opérateur"}
// ═══════════════════════════════════════════════════════════════
// 4. ACTION — cause fixe, sécurité d'abord, sans rotation
// Format (AF-07 §5.1) : [ORGANE] <Action physique> > <Fin>
// 🧊 Défauts (AU/puissance/SafeStop) + interlock DirectionBlocked
//    → affichés immédiatement (ForceInstant=TRUE) ; les autres états
//    → maintenus min (anti-clignotement).
// ═══════════════════════════════════════════════════════════════
IF CurrentMode = E_Mode.SEMI_AUTO THEN
    CurrentDirection := CycleRequestDirection;
ELSIF BothAxesCoupled THEN
    CurrentDirection := WinchBothMotionDirection;
ELSIF WinchSelected = 1 THEN
    CurrentDirection := M1LogicRequestDirection;
ELSIF WinchSelected = 2 THEN
    CurrentDirection := M2LogicRequestDirection;
ELSE
    CurrentDirection := 0;
END_IF;

DirectionBlocked := (CurrentDirection < 0 AND NOT DescendPermit)
                OR (CurrentDirection > 0 AND NOT AscentPermit);

// 🩹 Signaler la cause du dernier abandon de séquence AU (message cause+action),
// sans modifier le comportement de l'AU. Front descendant ArmingSeqStep (sequence en
// cours -> 0) = fin de sequence.
// 🐛 BUG A corrigé : l'ancien gating `NOT PowerContactorEngaged` supprimait le message
// d'abandon à l'étape 5 (PowerCutOff) car le contacteur venait d'être pulsé
// (PowerContactorEngaged=TRUE). On déclenche désormais sur la CAUSE (LastAbortCause <> 0),
// en excluant uniquement le SUCCÈS réel (séquence ayant atteint l'étape 6 de confirmation
// ET contacteur engagé au retour à IDLE) — un succès ne produit AUCUN message (AC4).
// Verrouillage : les causes SANS latch (CST_ABORT_POWER_CUTOFF, CST_ABORT_TIMEOUT_RESTORE_A/B)
// restauration) restent affichées jusqu'à Reset (ou nouvelle séquence) pour que
// l'opérateur voie l'échec. Les causes déjà latched (CST_ABORT_CHAIN_DROP/REDUNDANCY_A/B/
// TIMEOUT_CONTACTOR) et la coupe volontaire (CST_ABORT_CUT_IHM) ne sont pas verrouillées.
ArmingInProgress := (ArmingSeqStep <> 0);
LastAbortEdge(CLK := ArmingInProgress);
ResetEdge(CLK := Reset);
ArmStartEdge(CLK := ArmingInProgress);

// 🩹 Détection d'un SUCCÈS de séquence : la séquence a atteint l'étape 6 (confirmation).
// Ce drapeau est consommé par le test de LastAbortEdge ci-dessous AVANT d'être remis à
// zéro hors séquence (fin de bloc), pour distinguer un succès d'un abandon à l'étape 5.
IF ArmingSeqStep = 6 THEN
    SeqReachedConfirm := TRUE;
END_IF;

IF LastAbortEdge.Q AND (LastAbortCause <> 0) AND NOT (SeqReachedConfirm AND PowerContactorEngaged) THEN
    AbortMsgActive := TRUE;
    AbortMsgLatched := (LastAbortCause = INT_TO_WORD(CST_ABORT_POWER_CUTOFF)) OR (LastAbortCause = INT_TO_WORD(CST_ABORT_TIMEOUT_RESTORE_A)) OR (LastAbortCause = INT_TO_WORD(CST_ABORT_TIMEOUT_RESTORE_B));
    TonAbortHold(IN := FALSE);
END_IF;

// Effacement : Reset OU nouvelle séquence (évite le message périmé après réarmement réussi)
IF ResetEdge.Q OR ArmStartEdge.Q THEN
    AbortMsgActive := FALSE;
    AbortMsgLatched := FALSE;
    TonAbortHold(IN := FALSE);
END_IF;

// Remise à zéro du drapeau de confirmation hors séquence (après le test de LastAbortEdge
// ci-dessus, qui consomme sa valeur du scan précédent pour distinguer succès/abandon).
IF NOT ArmingInProgress THEN
    SeqReachedConfirm := FALSE;
END_IF;

// Maintien transitoire 5s UNIQUEMENT pour les causes non latched
IF AbortMsgActive AND NOT AbortMsgLatched THEN
    TonAbortHold(IN := TRUE, PT := CST_AbortHoldTime);
    IF TonAbortHold.Q THEN
        AbortMsgActive := FALSE;
        TonAbortHold(IN := FALSE);
    END_IF;
END_IF;
IF AbortMsgActive THEN
    IF LastAbortCause = INT_TO_WORD(CST_ABORT_CUT_IHM) THEN
        AbortMsgText := '[AU] Coupure volontaire IHM - relacher le bouton puis rearmer';
    ELSIF LastAbortCause = INT_TO_WORD(CST_ABORT_CHAIN_DROP) THEN
        AbortMsgText := '[AU] Boucle urgence ouverte (test) - relacher puis rearmer';
    ELSIF LastAbortCause = INT_TO_WORD(CST_ABORT_TIMEOUT_RESTORE_A) THEN
        AbortMsgText := '[AU] Chaine non remontee apres test A - verifier puis rearmer';
    ELSIF LastAbortCause = INT_TO_WORD(CST_ABORT_TIMEOUT_RESTORE_B) THEN
        AbortMsgText := '[AU] Chaine non remontee apres test B - verifier puis rearmer';
    ELSIF LastAbortCause = INT_TO_WORD(CST_ABORT_POWER_CUTOFF) THEN
        // 🩹 Décodage de la cause CST_ABORT_POWER_CUTOFF (PowerCutOff métier) en cause explicite
        // M1/M2/M3 + bit MecaA/MecaB/thermique, à partir des DUT Safety déjà en entrée.
        // Priorité : M3 (translation) puis M1 puis M2 ; MecaA > MecaB > thermique.
        IF TranslationSafety.ErrorMecaA THEN
            AbortMsgText := '[M3] MecaA (mouvement non commandé) - Reset puis réarmer';
        ELSIF TranslationSafety.ErrorMecaB THEN
            AbortMsgText := '[M3] MecaB (arrêt non confirmé) - Reset puis réarmer';
        ELSIF TranslationSafety.ErrorBrakeThermal THEN
            AbortMsgText := '[M3] Surchauffe frein - Reset puis réarmer';
        ELSIF WinchM1Safety.ErrorMecaA THEN
            AbortMsgText := '[M1] MecaA (mouvement non commandé) - Reset puis réarmer';
        ELSIF WinchM1Safety.ErrorMecaB THEN
            AbortMsgText := '[M1] MecaB (arrêt non confirmé) - Reset puis réarmer';
        ELSIF WinchM1Safety.ThermalFault THEN
            AbortMsgText := '[M1] Surchauffe moteur - Reset puis réarmer';
        ELSIF WinchM1Safety.ErrorBrakeThermal THEN
            AbortMsgText := '[M1] Surchauffe frein - Reset puis réarmer';
        ELSIF WinchM2Safety.ErrorMecaA THEN
            AbortMsgText := '[M2] MecaA (mouvement non commandé) - Reset puis réarmer';
        ELSIF WinchM2Safety.ErrorMecaB THEN
            AbortMsgText := '[M2] MecaB (arrêt non confirmé) - Reset puis réarmer';
        ELSIF WinchM2Safety.ThermalFault THEN
            AbortMsgText := '[M2] Surchauffe moteur - Reset puis réarmer';
        ELSIF WinchM2Safety.ErrorBrakeThermal THEN
            AbortMsgText := '[M2] Surchauffe frein - Reset puis réarmer';
        ELSE
            AbortMsgText := '[AU] Coupure securite metier active - lever la cause puis rearmer';
        END_IF;
    ELSIF LastAbortCause = INT_TO_WORD(CST_ABORT_REDUNDANCY_A) THEN
        AbortMsgText := '[AU] Defaut redondance canal A - verifier contacteur puis Reset';
    ELSIF LastAbortCause = INT_TO_WORD(CST_ABORT_REDUNDANCY_B) THEN
        AbortMsgText := '[AU] Defaut redondance canal B - verifier contacteur puis Reset';
    ELSIF LastAbortCause = INT_TO_WORD(CST_ABORT_TIMEOUT_CONTACTOR) THEN
        AbortMsgText := '[AU] Contacteur non engage sous 2s - verifier puis rearmer';
    ELSE
        AbortMsgText := '[AU] Rearmement interrompu - verifier et rearmer';
    END_IF;
END_IF;

// ═══════════════════════════════════════════════════════════════
// 🧊 MESSAGE DE REPLI AX_STAB — CAUSE RACINE (étape + cause cycle + cause winch)
// Construit AVANT la chaîne de priorités qui suit : toutes les causes winch décodables
// (MecaA/B/C/D/E, codeur, com opérateur, sens opposé, absence mouvement) SONT des causes
// SafeStop/PowerCutOff (FB_Safety_Winch §Agrégats) et restent vraies tant que le latch est
// posé. Sans cette priorité, le bandeau n'afficherait que « Acquitter SafeStop » ou
// « Coupure puissance » — conséquences, jamais la cause.
// ═══════════════════════════════════════════════════════════════
// CycleFaultActive et StepAtErrorStr sont calcules en §1bis (avant §2 et §4).
CycleFaultMsgStr := '';
IF CycleFaultActive THEN
    // Décodage priorisé de la cause cycle : l'opérateur voit la grandeur fautive, pas un masque.
    // Bits cycle : 0 limite, 1 synchro, 2 vitesse, 3 IHM, 4 tempo,
    // 5 stabilisation, 6 position, 7 FDC haut, 8/9 paliers, 10 arrêt.
    IF (CycleErrorId AND 16#0001) <> 0 THEN
        CycleFaultCauseStr := 'limite profondeur';
    ELSIF (CycleErrorId AND 16#0002) <> 0 THEN
        CycleFaultCauseStr := 'synchro M1/M2';
    ELSIF (CycleErrorId AND 16#0004) <> 0 THEN
        CycleFaultCauseStr := 'ecart vitesse M1/M2';
    ELSIF (CycleErrorId AND 16#0008) <> 0 THEN
        CycleFaultCauseStr := 'com IHM perdue';
    ELSIF (CycleErrorId AND 16#0010) <> 0 THEN
        CycleFaultCauseStr := 'tempo etape';
    ELSIF (CycleErrorId AND 16#0020) <> 0 THEN
        CycleFaultCauseStr := 'ecart codeurs remontee';
    ELSIF (CycleErrorId AND 16#0040) <> 0 THEN
        CycleFaultCauseStr := 'ecart position M1/M2';
    ELSIF (CycleErrorId AND 16#0080) <> 0 THEN
        CycleFaultCauseStr := 'hors FDC haut';
    ELSIF (CycleErrorId AND 16#0100) <> 0 THEN
        CycleFaultCauseStr := 'palier 5 interdit';
    ELSIF (CycleErrorId AND 16#0200) <> 0 THEN
        CycleFaultCauseStr := 'palier 4 non confirme';
    ELSIF (CycleErrorId AND 16#0400) <> 0 THEN
        CycleFaultCauseStr := 'arret meca non confirme';
    ELSIF (CycleErrorId AND 16#0800) <> 0 THEN
        CycleFaultCauseStr := 'consigne profondeur invalide';
    ELSE
        CycleFaultCauseStr := CONCAT('cause inconnue #', WORD_TO_STRING(CycleErrorId));
    END_IF;
    // 🔎 CAUSE RACINE WINCH — vue LATCHÉE (WinchMxSafety.LatchedId), jamais les bits LIVE : en
    // repli AX_STAB le cycle neutralise les ordres, donc le défaut safety live s'efface et
    // n'expliquerait plus rien. La vue latchée persiste jusqu'au Reset (acquittement).
    // Décodage PAR TREUIL : le masque et l'étiquette proviennent du MÊME treuil (M1 prioritaire),
    // pour ne jamais afficher la cause d'un treuil avec l'étiquette de l'autre (multi-latch).
    WinchRootCauseStr := '';
    WinchRootCauseLbl := '';
    WinchRootTagStr   := '';
    WinchRootMaskId   := 0;
    IF WinchM1Safety.LatchedId <> 0 THEN
        WinchRootTagStr := 'M1 ';
        WinchRootMaskId := WinchM1Safety.LatchedId;
    ELSIF WinchM2Safety.LatchedId <> 0 THEN
        WinchRootTagStr := 'M2 ';
        WinchRootMaskId := WinchM2Safety.LatchedId;
    END_IF;
    IF WinchRootMaskId <> 0 THEN
        IF (WinchRootMaskId AND 16#3000) <> 0 THEN
            WinchRootCauseLbl := 'MecaE';
        ELSIF (WinchRootMaskId AND 16#0080) <> 0 THEN
            WinchRootCauseLbl := 'MecaA';
        ELSIF (WinchRootMaskId AND 16#0100) <> 0 THEN
            WinchRootCauseLbl := 'MecaB';
        ELSIF (WinchRootMaskId AND 16#0200) <> 0 THEN
            WinchRootCauseLbl := 'MecaC';
        ELSIF (WinchRootMaskId AND 16#0800) <> 0 THEN
            WinchRootCauseLbl := 'MecaD';
        ELSIF (WinchRootMaskId AND 16#0002) <> 0 THEN
            WinchRootCauseLbl := 'codeur';
        ELSIF (WinchRootMaskId AND 16#0001) <> 0 THEN
            WinchRootCauseLbl := 'com op';
        ELSIF (WinchRootMaskId AND 16#4000) <> 0 THEN
            WinchRootCauseLbl := 'sens opp';
        ELSIF (WinchRootMaskId AND 16#8000) <> 0 THEN
            WinchRootCauseLbl := 'sans mvt';
        END_IF;
    END_IF;
    // Mou de câble : vue LIVE seule (non latchée dans FB_Safety_Winch) — sans étiquette treuil
    // car la détection est commune M1/M2 (les deux lisent M2_TensionedCable_DI).
    IF WinchRootMaskId = 0 THEN
        IF WinchM1Safety.SlackCable OR WinchM2Safety.SlackCable THEN
            WinchRootCauseLbl := 'mou cable';
            WinchRootTagStr   := '';
        END_IF;
    END_IF;
    IF WinchRootCauseLbl <> '' THEN
        WinchRootCauseStr := CONCAT(' (', CONCAT(WinchRootTagStr,
                                 CONCAT(WinchRootCauseLbl, ')')));
    END_IF;
    // Concaténation (jamais substitution) : cause dérivée cycle PUIS cause racine.
    CycleFaultMsgStr := CONCAT('[CYCLE]', CONCAT(StepAtErrorStr,
                        CONCAT(':', CONCAT(CycleFaultCauseStr,
                        CONCAT(WinchRootCauseStr, '>Repr/Abandon')))));
END_IF;

IF NOT EmergencyChainClosed THEN
    OperatorActionCandidate := '[PUPITRE] Boucle urgence ouverte - réarmer';
ELSIF NOT LocalIoValid OR NOT Vh0800Valid OR NOT Vh0808Valid OR NOT Vh0008ErValid OR NOT Vh0008Er1Valid THEN
    OperatorActionCandidate := '[IO] Défaut module E/S - vérifier alimentation/coupleur';
ELSIF NOT CanBusValid THEN
    OperatorActionCandidate := '[CAN] Défaut bus CANopen - vérifier câblage';
ELSIF NOT Joy1Valid THEN
    OperatorActionCandidate := '[CAN] Joystick non détecté - vérifier liaison';
ELSIF NOT EcatBusValid THEN
    OperatorActionCandidate := '[ECAT] Défaut bus EtherCAT - vérifier liaison';
ELSIF NOT EncM1Valid OR NOT EncM2Valid THEN
    OperatorActionCandidate := '[ECAT] Codeurs non détectés - vérifier liaison';
ELSIF NOT VarM3Valid THEN
    OperatorActionCandidate := '[ECAT] Variateur non détecté - vérifier liaison';
ELSIF AbortMsgActive THEN
    // 🩹 Cause du dernier abandon de séquence AU (message explicite cause+action).
    // 🐛 BUG B corrigé : placé AVANT PowerCutOffActiveAny pour que la cause racine
    // (dont CST_ABORT_POWER_CUTOFF décodée en M1/M2/M3 + MecaA/MecaB/thermique) prime sur
    // le message générique de coupure puissance. Placé aussi avant
    // RedundancyTestFailed/EmergencyArmingFailed/SafeStop pour que chaque cause montre
    // son message spécifique — le message d'abandon est la CAUSE RACINE (plus pertinente
    // que le SafeStop qui en est une conséquence) — il prime sur SafeStop/DirectionBlocked.
    OperatorActionCandidate := AbortMsgText;
ELSIF CycleFaultActive THEN
    // 🩹 Repli AX_STAB sur défaut cycle : la CAUSE RACINE (étape d'origine + cause cycle +
    // cause winch latchée) PRIME sur les messages génériques de coupure puissance et de
    // SafeStop, qui n'en sont que la CONSÉQUENCE (toutes les causes winch Meca* sont des
    // causes SafeStop/PowerCutOff et resteraient affichées sinon).
    OperatorActionCandidate := CycleFaultMsgStr;
ELSIF PowerCutOffActiveAny THEN
    OperatorActionCandidate := '[SÉCURITÉ] Coupure puissance active - acquitter défaut treuil/pont';
ELSIF RedundancyTestFailed THEN
    OperatorActionCandidate := '[AU] Défaut redondance contacteurs - réarmer (Reset)';
ELSIF EmergencyArmingFailed THEN
    OperatorActionCandidate := '[AU] Échec réarmement contacteur - réarmer';
ELSIF NOT PowerContactorEngaged THEN
    OperatorActionCandidate := '[PUPITRE] Réarmer AU et puissance';
ELSIF SafeStopActive THEN
    IF SyncContactorDiag.MismatchLevel >= 1 THEN
        OperatorActionCandidate := '[SYNC] Discordance contacteurs M1/M2 - Acquitter SafeStop';
    ELSIF WinchM1Safety.SlackCable OR WinchM2Safety.SlackCable THEN
        OperatorActionCandidate := '[TREUIL] Mou de cable detecte - retendre ou acquitter';
    ELSE
        OperatorActionCandidate := '[PUPITRE] Acquitter SafeStop';
    END_IF;
ELSIF DirectionBlocked THEN
    IF CurrentDirection < 0 THEN
        IF WinchDescentLockedByM3 THEN
            // 🛡️ Descente verrouillée par position M3 (chariot pas à P1/Maintenance)
            OperatorActionCandidate := '[TREUIL] Descente interdite - Chariot M3 pas a P1/Maintenance';
        ELSIF LegalLimitReached THEN
            // 🛡️ Descente bloquée par limite légale atteinte
            OperatorActionCandidate := '[TREUIL] Descente interdite - Limite legale atteinte';
        ELSIF WinchM1Safety.CableLimitDescent OR WinchM2Safety.CableLimitDescent THEN
            // 🛡️ Descente bloquée par limite basse câble
            OperatorActionCandidate := '[TREUIL] Descente interdite - Limite basse cable';
        ELSIF WinchM1Safety.SlackCable OR WinchM2Safety.SlackCable THEN
            // 🛡️ Descente bloquée par détection mou de câble
            OperatorActionCandidate := '[TREUIL] Descente interdite - Mou de cable detecte';
        ELSIF WinchM1Safety.DescendPermit AND NOT WinchM2Safety.DescendPermit THEN
            // 🛡️ Descente bloquée spécifiquement par M2
            OperatorActionCandidate := '[TREUIL] Descente interdite - Treuil M2 (benne)';
        ELSIF WinchM2Safety.DescendPermit AND NOT WinchM1Safety.DescendPermit THEN
            // 🛡️ Descente bloquée spécifiquement par M1
            OperatorActionCandidate := '[TREUIL] Descente interdite - Treuil M1 (retenue)';
        ELSE
            OperatorActionCandidate := '[TREUIL] Descente interdite';
        END_IF;
    ELSIF TopHardStopLatched THEN
        OperatorActionCandidate := 'Position haute deja depassee - redescendre pour degager';
    ELSIF TopPositionSensorActive THEN
        OperatorActionCandidate := '[TREUIL] Montee interdite - capteur haut';
    ELSIF TopLimitReached THEN
        // 🛡️ Montée bloquée par butée logicielle haute (agrégat M1/M2) — cause exposée par le safety.
        OperatorActionCandidate := '[TREUIL] Montée interdite - limite haute';
    ELSIF WinchM1Safety.ErrorMecaD OR WinchM2Safety.ErrorMecaD THEN
        // 🛡️ Montée bloquée par capteur haut (non-arrêt au capteur haut, MecaD) — cause exposée par le safety.
        OperatorActionCandidate := '[TREUIL] Montée interdite - capteur haut';
    ELSIF WinchM1Safety.AscentPermit AND NOT WinchM2Safety.AscentPermit THEN
        // 🛡️ Montée bloquée par treuil M2 (M1 autorise, M2 non) — cause exposée par le safety.
        OperatorActionCandidate := '[TREUIL] Montée interdite - treuil M2';
    ELSE
        OperatorActionCandidate := '[TREUIL] Montée interdite';
    END_IF;
ELSIF CfgCorrectedT330 THEN
    // 🔧 T330 — reglage haut corrige automatiquement (Q2). Volontairement place APRES toutes
    // les branches de SECURITE (AU, puissance, SafeStop, direction) : une correction de reglage
    // ne doit JAMAIS masquer une alarme de securite. Prefixe [CFG] discriminant pour rester
    // distinguable de D18, benne non fermee et synchro (cadrage §11bis). Longueur <= 70 car. (G408).
    OperatorActionCandidate := '[CFG] Reglage corrige : reserve TOP/FDC a 1,00 m';
ELSIF CurrentMode = E_Mode.DISABLE THEN
    OperatorActionCandidate := '[IHM] Sélectionner un mode';
ELSIF TopHardStopLatched AND NOT MachineHomingActive THEN
    OperatorActionCandidate := 'Position haute deja depassee - redescendre pour degager';
ELSIF (MachineHomingActive OR MachineHomingFailed
       OR ((CurrentMode = E_Mode.MAINT_N1) AND (MachineHomingStep > 0) AND (MachineHomingStep <> 60)))
      AND (MachineHomingActionText <> '') THEN
    // Consignes directes du GRAFCET homing : priment sur les actions generiques joystick/benne.
    OperatorActionCandidate := MachineHomingActionText;
ELSIF CurrentMode = E_Mode.SEMI_AUTO THEN
    // Guidance par étape du cycle (AF-07 §5.1) — ne masque jamais un défaut
    // (priorités AU/puissance/SafeStop/DirectionBlocked ci-dessus dominent).
    CASE CycleStep OF
        E_AutoCycleStep.AX0_REPOS:
            OperatorActionCandidate := '[IHM-JOY] Appuyer Start Cycle (ou homme-mort) pour initialiser';
        E_AutoCycleStep.AX1_INIT:
            IF CycleStateStr <> '' THEN
                OperatorActionCandidate := CONCAT('[INIT] ', CycleStateStr);
            ELSE
                OperatorActionCandidate := '[INIT] Verifier conditions initiales (referencement, FDC haut)';
            END_IF;
        E_AutoCycleStep.AX2_TRANSLATE_P1:
            OperatorActionCandidate := '[JOY] Pousser a droite : translation vers P1';
        E_AutoCycleStep.AX3_OPEN_BUCKET:
            OperatorActionCandidate := '[JOY] Pousser descente : ouverture benne jusqu au FDC';
        E_AutoCycleStep.AX4_DESCEND_DIVING:
            OperatorActionCandidate := '[JOY] Pousser descente : plongee palier 4';
        E_AutoCycleStep.AX5_KOBOLD_INIT:
            OperatorActionCandidate := '[JOY] Maintenir descente : init Kobold';
        E_AutoCycleStep.AX6_SEARCH_IMMERSION:
            OperatorActionCandidate := '[JOY] Maintenir descente : recherche immersion';
        E_AutoCycleStep.AX7_SEARCH_BOTTOM:
            OperatorActionCandidate := '[JOY] Maintenir descente : recherche fond (Kobold)';
        E_AutoCycleStep.AX8_BOTTOM_CONFIRMED:
            OperatorActionCandidate := '[JOY] Fond atteint : relacher puis tirer pour extraire';
        E_AutoCycleStep.AX_DIVING_RETRY:
            OperatorActionCandidate := '[JOY] Reprise plongee : remonter au FDC haut';
        E_AutoCycleStep.AX9_RAISE_OFF_BOTTOM:
            OperatorActionCandidate := '[JOY] Tirer : montee synchronisee et retendre les cables';
        E_AutoCycleStep.AX10_CLOSE_BUCKET:
            OperatorActionCandidate := '[JOY] Tirer montee : fermeture de la benne';
        E_AutoCycleStep.AX11_CTRL_ASCENT:
            OperatorActionCandidate := '[JOY] Tirer montee : remontee de controle';
        E_AutoCycleStep.AX12_LOADED_ASCENT:
            OperatorActionCandidate := '[JOY] Tirer montee : remontee en charge';
        E_AutoCycleStep.AX13_DRAIN_PAUSE:
            OperatorActionCandidate := '[CYCLE] Egouttage en cours (attendre tempo ou bouton Passer)';
        E_AutoCycleStep.AX14_TRANSLATE_DUMP:
            OperatorActionCandidate := '[JOY] Pousser a gauche : translation vers tremie';
        E_AutoCycleStep.AX15A_DUMP_ARRIVE, E_AutoCycleStep.AX15B_DUMP_OPEN:
            OperatorActionCandidate := '[JOY] Pousser descente : vidage benne a la tremie';
        E_AutoCycleStep.AX15C_DUMP_REPOSITION:
            OperatorActionCandidate := '[JOY] Pousser descente : vidage benne a la tremie';
        E_AutoCycleStep.AX18_DONE_SYNC:
            OperatorActionCandidate := '[JOY] Cycle termine : pousser a droite vers P1';
        E_AutoCycleStep.AX_STAB:
            // Repli défaut : le message complet (étape d'origine + cause cycle + cause racine
            // winch) est construit AVANT la chaîne de priorités, pour que la CAUSE prime sur les
            // messages génériques SafeStop / coupure puissance qui n'en sont que la conséquence.
            OperatorActionCandidate := CycleFaultMsgStr;
        ELSE
            OperatorActionCandidate := '[CYCLE] Cycle en cours...';
    END_CASE;
ELSIF DiveActive AND CurrentDirection < 0 THEN
    OperatorActionCandidate := '[TREUIL] Attendre fin du Dive';
ELSIF NOT BucketIsOpen AND CurrentDirection < 0 THEN
    OperatorActionCandidate := '[BENNE] Ouvrir la benne';
ELSIF TopLimitReached AND CurrentDirection > 0 THEN
    OperatorActionCandidate := '[TREUIL] Limite haute';
ELSIF NOT BucketIsClosed AND CurrentDirection > 0 THEN
    // Sécurité : benne mal fermée (branche/caillou) → montee bridee palier 1 pour eviter un choc
    // si la benne se refermait d'un coup en montant vite.
    OperatorActionCandidate := '[BENNE] Benne non fermee - montee bridee palier 1 (securite)';
ELSIF CurrentMode = E_Mode.DISABLE THEN
    OperatorActionCandidate := '[IHM] Sélectionner un mode';
ELSIF ArmingPermitDenied THEN
    CASE ArmingBlockedReason OF
        E_ArmingBlockReason.MODE_DISABLE:
            OperatorActionCandidate := '[JOYSTICK] Armement refusé : mode DÉSACTIVÉ';
        E_ArmingBlockReason.CONTACTOR_OFF:
            OperatorActionCandidate := '[JOYSTICK] Armement refusé : contacteur puissance non enclenché';
        E_ArmingBlockReason.POWER_CUTOFF:
            OperatorActionCandidate := '[JOYSTICK] Armement refusé : coupure puissance active';
        E_ArmingBlockReason.BUCKET_BUSY:
            OperatorActionCandidate := '[JOYSTICK] Armement refusé : action benne en cours';
        E_ArmingBlockReason.ALL_AXES_BLOCKED:
            OperatorActionCandidate := '[JOYSTICK] Armement refusé : aucun axe disponible';
    ELSE
        OperatorActionCandidate := '[JOYSTICK] Armement refusé : mouvements non autorisés';
    END_CASE;
ELSIF TopHardStopLatched THEN
    OperatorActionCandidate := 'Position haute deja depassee - redescendre pour degager';
ELSIF NOT DeadmanArmed THEN
    OperatorActionCandidate := '[JOYSTICK] Appuyer homme-mort au neutre';
ELSIF ((WinchM1Safety.ErrorId OR WinchM2Safety.ErrorId) AND CST_WinchErrorIdCableLimitDescent) <> 16#0000 THEN
    // 🛡️ Cause limite basse câble ACTIVE (bit 6) ⇒ descente INTERDITE
    // (DescendPermit = FALSE, FB_Safety_Winch.st:563-565) et REMONTÉE = seule action
    // autorisée. Nomme la cause ET l'action même SANS commande de descente : la branche
    // « Descente interdite - Limite basse cable » (ligne 661) n'est atteinte que si
    // DirectionBlocked = TRUE, donc jamais joystick relâché.
    // Lue sur ErrorId (cause safety, bypass et mode référencement respectés) et jamais sur
    // WinchMxSafety.CableLimitDescent, champ de projection brute sans bypass.
    // Ordre volontaire : APRÈS « Descente interdite » (une descente réellement commandée
    // garde son libellé historique) et APRÈS la branche DISABLE (aucune action proposée
    // hors mode de marche), AVANT les rappels joystick : la cause prime sur le guidage,
    // jamais sur un prérequis de mode.
    IF ((WinchM1Safety.ErrorId AND WinchM2Safety.ErrorId) AND CST_WinchErrorIdCableLimitDescent) <> 16#0000 THEN
        OperatorActionCandidate := '[TREUIL] Limite basse cable M1+M2 - remonter';
    ELSIF (WinchM1Safety.ErrorId AND CST_WinchErrorIdCableLimitDescent) <> 16#0000 THEN
        OperatorActionCandidate := '[TREUIL] Limite basse cable M1 - remonter';
    ELSE
        OperatorActionCandidate := '[TREUIL] Limite basse cable M2 - remonter';
    END_IF;
ELSIF JoystickAtNeutral THEN
    OperatorActionCandidate := '[JOYSTICK] Armé - actionner axe';
ELSE
    OperatorActionCandidate := '[JOYSTICK] Déplacement en cours';
END_IF;

// Interlock = mouvement demandé mais permit absent : c'est une cause
// sécurité (blocage de mouvement) → affichage IMMÉDIAT, comme un défaut.
PowerOrChainFault := (NOT EmergencyChainClosed OR NOT PowerContactorEngaged OR PowerCutOffActiveAny);
HardwareModuleOrBusFault := (NOT LocalIoValid OR NOT Vh0800Valid OR NOT Vh0808Valid OR NOT Vh0008ErValid OR NOT Vh0008Er1Valid OR NOT CanBusValid OR NOT Joy1Valid OR NOT EcatBusValid OR NOT EncM1Valid OR NOT EncM2Valid OR NOT VarM3Valid);
CriticalActionActive := (PowerOrChainFault OR HardwareModuleOrBusFault OR SafeStopActive OR DirectionBlocked OR ArmingPermitDenied OR TopHardStopLatched OR CycleFaultActive OR MachineHomingActive OR MachineHomingFailed);

AntiFlickOperator(NewText := OperatorActionCandidate, ForceInstant := CriticalActionActive, HoldTime := CST_BannerHoldTime);
Banner.OperatorActionText := AntiFlickOperator.Text;
{endregion}

{region "§5 Bandeau alarme"}
// ═══════════════════════════════════════════════════════════════
// 5. BANDEAU D'ALARME — carrousel des défauts actifs (index n/N)
// Format (AF-07 §6) : [ORGANE] raison_brève. Un défaut à la fois,
// rotation 1→2→…→N→1, maintien AlarmHoldTime par message.
// 🧊 Distinct des 4 champs ci-dessus (AF-07 §5.2) : ce carrousel est
//    le SEUL endroit du bandeau qui publie Error/ErrorId (alarmes).
// ═══════════════════════════════════════════════════════════════
AlarmCount := 0;

// 5.0 Collecte — Défauts matériels parents (priorité absolue carrousel)
IF NOT LocalIoValid AND (AlarmCount < CST_NbMaxAlarmes) THEN
    AlarmArray[AlarmCount] := '[IO] Defaut module Local IO (DI8/DO8)'; AlarmCount := AlarmCount + 1;
END_IF;
IF NOT Vh0800Valid AND (AlarmCount < CST_NbMaxAlarmes) THEN
    AlarmArray[AlarmCount] := '[IO] Defaut module VH0800END (DI8)'; AlarmCount := AlarmCount + 1;
END_IF;
IF NOT Vh0808Valid AND (AlarmCount < CST_NbMaxAlarmes) THEN
    AlarmArray[AlarmCount] := '[IO] Defaut module VH0808ETP (DI8/DO8)'; AlarmCount := AlarmCount + 1;
END_IF;
IF NOT Vh0008ErValid AND (AlarmCount < CST_NbMaxAlarmes) THEN
    AlarmArray[AlarmCount] := '[IO] Defaut module VH0008ER (DO8 Relais)'; AlarmCount := AlarmCount + 1;
END_IF;
IF NOT Vh0008Er1Valid AND (AlarmCount < CST_NbMaxAlarmes) THEN
    AlarmArray[AlarmCount] := '[IO] Defaut module VH0008ER_1 (DO8 Relais)'; AlarmCount := AlarmCount + 1;
END_IF;
IF NOT CanBusValid AND (AlarmCount < CST_NbMaxAlarmes) THEN
    AlarmArray[AlarmCount] := '[CAN] Defaut bus CANopen'; AlarmCount := AlarmCount + 1;
END_IF;
IF CanBusValid AND NOT Joy1Valid AND (AlarmCount < CST_NbMaxAlarmes) THEN
    AlarmArray[AlarmCount] := '[CAN] Joystick JOY1 non detecte'; AlarmCount := AlarmCount + 1;
END_IF;
IF NOT EcatBusValid AND (AlarmCount < CST_NbMaxAlarmes) THEN
    AlarmArray[AlarmCount] := '[ECAT] Defaut bus EtherCAT'; AlarmCount := AlarmCount + 1;
END_IF;
IF NOT EncM1Valid AND (AlarmCount < CST_NbMaxAlarmes) THEN
    AlarmArray[AlarmCount] := '[M1] Codeur absolu COD1 non detecte (ECAT)'; AlarmCount := AlarmCount + 1;
END_IF;
IF NOT EncM2Valid AND (AlarmCount < CST_NbMaxAlarmes) THEN
    AlarmArray[AlarmCount] := '[M2] Codeur absolu COD2 non detecte (ECAT)'; AlarmCount := AlarmCount + 1;
END_IF;
IF NOT VarM3Valid AND (AlarmCount < CST_NbMaxAlarmes) THEN
    AlarmArray[AlarmCount] := '[M3] Variateur AC600 non detecte (ECAT)'; AlarmCount := AlarmCount + 1;
END_IF;

// 5a. Collecte — treuil M1 (ST_SafetyWinch, bits ErrorId décodés)
// 🧊 Tri bloquant/warning (AF-07 §6, décision 2026-09-01) : seuls les défauts
//    BLOQUANTS (SafeStop/PowerCutOff/interlock) sont publiés. Les warnings non
//    bloquants (mou de câble, surchauffe moteur/frein, limites basse/haute) sont
//    EXCLUS du carrousel — ils restent visibles via OperatorActionText/SpecialCondition.
IF WinchM1Safety.ErrorOperatorComm AND Joy1Valid AND (AlarmCount < CST_NbMaxAlarmes) THEN
    AlarmArray[AlarmCount] := '[M1] ErrorID:01 - perte com operateur'; AlarmCount := AlarmCount + 1;
END_IF;
IF WinchM1Safety.ErrorEncoder AND (AlarmCount < CST_NbMaxAlarmes) THEN
    AlarmArray[AlarmCount] := '[M1] ErrorID:02 - perte codeur'; AlarmCount := AlarmCount + 1;
END_IF;
IF WinchM1Safety.ThermalFault AND (AlarmCount < CST_NbMaxAlarmes) THEN
    AlarmArray[AlarmCount] := '[M1] ErrorID:03 - surchauffe moteur'; AlarmCount := AlarmCount + 1;
END_IF;
IF WinchM1Safety.ErrorPhaseRotation AND Vh0800Valid AND (AlarmCount < CST_NbMaxAlarmes) THEN
    AlarmArray[AlarmCount] := '[M1] ErrorID:05 - rotation phases'; AlarmCount := AlarmCount + 1;
END_IF;
IF WinchM1Safety.ErrorMecaA AND EncM1Valid AND (AlarmCount < CST_NbMaxAlarmes) THEN
    AlarmArray[AlarmCount] := '[M1] ErrorID:08 - MecaA - deplacement sans commande'; AlarmCount := AlarmCount + 1;
END_IF;
IF WinchM1Safety.ErrorMecaB AND EncM1Valid AND (AlarmCount < CST_NbMaxAlarmes) THEN
    AlarmArray[AlarmCount] := '[M1] ErrorID:09 - MecaB - arret non confirme apres stop'; AlarmCount := AlarmCount + 1;
END_IF;
IF WinchM1Safety.ErrorMecaC AND EncM1Valid AND EncM2Valid AND (AlarmCount < CST_NbMaxAlarmes) THEN
    AlarmArray[AlarmCount] := '[M1] ErrorID:10 - MecaC - glissement pendant benne figee'; AlarmCount := AlarmCount + 1;
END_IF;
IF WinchM1Safety.ErrorBrakeThermal AND (AlarmCount < CST_NbMaxAlarmes) THEN
    AlarmArray[AlarmCount] := '[M1] ErrorID:11 - surchauffe frein'; AlarmCount := AlarmCount + 1;
END_IF;
IF WinchM1Safety.ErrorMecaD AND LocalIoValid AND EncM1Valid AND (AlarmCount < CST_NbMaxAlarmes) THEN
    AlarmArray[AlarmCount] := '[M1] ErrorID:12 - MecaD - non-arret au capteur haut'; AlarmCount := AlarmCount + 1;
END_IF;
IF WinchM1Safety.ErrorMecaE AND EncM1Valid AND EncM2Valid AND (AlarmCount < CST_NbMaxAlarmes) THEN
    AlarmArray[AlarmCount] := '[M1] ErrorID:13 - MecaE - ecart synchro M1/M2 critique'; AlarmCount := AlarmCount + 1;
END_IF;
IF WinchM1Safety.ErrorOppositeDir AND EncM1Valid AND (AlarmCount < CST_NbMaxAlarmes) THEN
    AlarmArray[AlarmCount] := '[M1] ErrorID:15 - sens oppose'; AlarmCount := AlarmCount + 1;
END_IF;
IF WinchM1Safety.ErrorNoMovement AND EncM1Valid AND (AlarmCount < CST_NbMaxAlarmes) THEN
    AlarmArray[AlarmCount] := '[M1] ErrorID:16 - discordance commande/retour/mouvement'; AlarmCount := AlarmCount + 1;
END_IF;
IF WinchM1Safety.ErrorOverspeed AND EncM1Valid AND (AlarmCount < CST_NbMaxAlarmes) THEN
    AlarmArray[AlarmCount] := '[M1] Survitesse treuil detectee (SafeStop)'; AlarmCount := AlarmCount + 1;
END_IF;
// 🛡️ 5a-bis. Limite de course BASSE du treuil M1 : cause BLOQUANTE (DescendPermit,
//    FB_Safety_Winch.st:563-565), donc publiée au carrousel au titre d'AF-07 §6 (interlock).
//    Cause 6 = instCauses[6].Active (FB_Safety_Winch.st:318-325), bit 6 = 16#0040, NON
//    latchée : elle allume AnyFaultActive via Safety.Error (PRG_07:541-542) et n'est
//    présente ni en vue active sans cette entrée, ni en [HISTO] (jamais dans LatchedId).
//    ⚠️ Lue sur ErrorId (la CAUSE safety, qui respecte tous les bypass) et JAMAIS sur
//    WinchM1Safety.CableLimitDescent, champ de projection brute sans bypass
//    (FB_WinchStateProjection.st:217-218/230) : le lire produirait une FAUSSE alarme sous
//    BypassCableLimitSwitch (MAINT_N2).
//    Gardée par la validité encodeur, comme les autres alarmes filles du treuil.
IF (WinchM1Safety.ErrorId AND CST_WinchErrorIdCableLimitDescent) <> 16#0000 AND EncM1Valid AND (AlarmCount < CST_NbMaxAlarmes) THEN
    AlarmArray[AlarmCount] := '[M1] Limite basse cable atteinte'; AlarmCount := AlarmCount + 1;
END_IF;

// 5b. Collecte — treuil M2 (mêmes bits que M1, tri bloquant/warning identique)
IF WinchM2Safety.ErrorOperatorComm AND Joy1Valid AND (AlarmCount < CST_NbMaxAlarmes) THEN
    AlarmArray[AlarmCount] := '[M2] ErrorID:01 - perte com operateur'; AlarmCount := AlarmCount + 1;
END_IF;
IF WinchM2Safety.ErrorEncoder AND (AlarmCount < CST_NbMaxAlarmes) THEN
    AlarmArray[AlarmCount] := '[M2] ErrorID:02 - perte codeur'; AlarmCount := AlarmCount + 1;
END_IF;
IF WinchM2Safety.ThermalFault AND (AlarmCount < CST_NbMaxAlarmes) THEN
    AlarmArray[AlarmCount] := '[M2] ErrorID:03 - surchauffe moteur'; AlarmCount := AlarmCount + 1;
END_IF;
IF WinchM2Safety.ErrorPhaseRotation AND Vh0800Valid AND (AlarmCount < CST_NbMaxAlarmes) THEN
    AlarmArray[AlarmCount] := '[M2] ErrorID:05 - rotation phases'; AlarmCount := AlarmCount + 1;
END_IF;
IF WinchM2Safety.ErrorMecaA AND EncM2Valid AND (AlarmCount < CST_NbMaxAlarmes) THEN
    AlarmArray[AlarmCount] := '[M2] ErrorID:08 - MecaA - deplacement sans commande'; AlarmCount := AlarmCount + 1;
END_IF;
IF WinchM2Safety.ErrorMecaB AND EncM2Valid AND (AlarmCount < CST_NbMaxAlarmes) THEN
    AlarmArray[AlarmCount] := '[M2] ErrorID:09 - MecaB - arret non confirme apres stop'; AlarmCount := AlarmCount + 1;
END_IF;
IF WinchM2Safety.ErrorMecaC AND EncM1Valid AND EncM2Valid AND (AlarmCount < CST_NbMaxAlarmes) THEN
    AlarmArray[AlarmCount] := '[M2] ErrorID:10 - MecaC - glissement pendant benne figee'; AlarmCount := AlarmCount + 1;
END_IF;
IF WinchM2Safety.ErrorBrakeThermal AND (AlarmCount < CST_NbMaxAlarmes) THEN
    AlarmArray[AlarmCount] := '[M2] ErrorID:11 - surchauffe frein'; AlarmCount := AlarmCount + 1;
END_IF;
IF WinchM2Safety.ErrorMecaD AND LocalIoValid AND EncM2Valid AND (AlarmCount < CST_NbMaxAlarmes) THEN
    AlarmArray[AlarmCount] := '[M2] ErrorID:12 - MecaD - non-arret au capteur haut'; AlarmCount := AlarmCount + 1;
END_IF;
IF WinchM2Safety.ErrorMecaE AND EncM1Valid AND EncM2Valid AND (AlarmCount < CST_NbMaxAlarmes) THEN
    AlarmArray[AlarmCount] := '[M2] ErrorID:13 - MecaE - ecart synchro M1/M2 critique'; AlarmCount := AlarmCount + 1;
END_IF;
IF WinchM2Safety.ErrorOppositeDir AND EncM2Valid AND (AlarmCount < CST_NbMaxAlarmes) THEN
    AlarmArray[AlarmCount] := '[M2] ErrorID:15 - sens oppose'; AlarmCount := AlarmCount + 1;
END_IF;
IF WinchM2Safety.ErrorNoMovement AND EncM2Valid AND (AlarmCount < CST_NbMaxAlarmes) THEN
    AlarmArray[AlarmCount] := '[M2] ErrorID:16 - discordance commande/retour/mouvement'; AlarmCount := AlarmCount + 1;
END_IF;
IF WinchM2Safety.ErrorOverspeed AND EncM2Valid AND (AlarmCount < CST_NbMaxAlarmes) THEN
    AlarmArray[AlarmCount] := '[M2] Survitesse treuil detectee (SafeStop)'; AlarmCount := AlarmCount + 1;
END_IF;
// 🛡️ 5b-bis. Limite de course BASSE du treuil M2 — même cause, mêmes raisons que 5a-bis.
IF (WinchM2Safety.ErrorId AND CST_WinchErrorIdCableLimitDescent) <> 16#0000 AND EncM2Valid AND (AlarmCount < CST_NbMaxAlarmes) THEN
    AlarmArray[AlarmCount] := '[M2] Limite basse cable atteinte'; AlarmCount := AlarmCount + 1;
END_IF;

// 5c. Collecte — translation M3 (ST_SafetyTranslation, tri bloquant/warning identique)
IF TranslationSafety.ErrorOperatorComm AND Joy1Valid AND (AlarmCount < CST_NbMaxAlarmes) THEN
    AlarmArray[AlarmCount] := '[M3] ErrorID:01 - perte com operateur'; AlarmCount := AlarmCount + 1;
END_IF;
IF TranslationSafety.ErrorDriveComm AND VarM3Valid AND (AlarmCount < CST_NbMaxAlarmes) THEN
    AlarmArray[AlarmCount] := '[M3] ErrorID:02 - perte EtherCAT'; AlarmCount := AlarmCount + 1;
END_IF;
IF TranslationSafety.ErrorPhaseRotation AND Vh0800Valid AND (AlarmCount < CST_NbMaxAlarmes) THEN
    AlarmArray[AlarmCount] := '[M3] ErrorID:03 - rotation phases'; AlarmCount := AlarmCount + 1;
END_IF;
IF TranslationSafety.ErrorBrakeThermal AND (AlarmCount < CST_NbMaxAlarmes) THEN
    AlarmArray[AlarmCount] := '[M3] ErrorID:04 - surchauffe frein'; AlarmCount := AlarmCount + 1;
END_IF;
IF TranslationSafety.ErrorMecaB AND VarM3Valid AND (AlarmCount < CST_NbMaxAlarmes) THEN
    AlarmArray[AlarmCount] := '[M3] ErrorID:05 - MecaB - arret non confirme apres stop'; AlarmCount := AlarmCount + 1;
END_IF;
IF TranslationSafety.ErrorMecaA AND VarM3Valid AND (AlarmCount < CST_NbMaxAlarmes) THEN
    AlarmArray[AlarmCount] := '[M3] ErrorID:06 - MecaA - deplacement sans commande'; AlarmCount := AlarmCount + 1;
END_IF;
IF TranslationSafety.ErrorLimitSwitch AND Vh0808Valid AND (AlarmCount < CST_NbMaxAlarmes) THEN
    AlarmArray[AlarmCount] := '[M3] ErrorID:07 - butee extreme'; AlarmCount := AlarmCount + 1;
END_IF;
IF TranslationSafety.ErrorSensorIncoherent AND Vh0808Valid AND (AlarmCount < CST_NbMaxAlarmes) THEN
    AlarmArray[AlarmCount] := '[M3] ErrorID:08 - capteurs incoherents'; AlarmCount := AlarmCount + 1;
END_IF;
// 5c-bis. Defauts MOUVEMENT M3 (FB_Translation.Fault) — distincts des defauts SAFETY
//    ci-dessus. Ils n'avaient AUCUN chemin vers le carrousel d'alarmes (regression MES
//    2026-09-04 : "M3 chariot fault" invisible). Bits FB_FaultCore : 0=frein, 3=variateur
//    AC600 (latching), 6=limite extreme. + barriere finale (frein/redemarrage).
IF ((TranslationMotionErrorId AND 16#0001) <> 16#0000) AND (AlarmCount < CST_NbMaxAlarmes) THEN
    AlarmArray[AlarmCount] := '[M3] Defaut sequence / retour frein translation'; AlarmCount := AlarmCount + 1;
END_IF;
IF ((TranslationMotionErrorId AND 16#0008) <> 16#0000) AND VarM3Valid AND (AlarmCount < CST_NbMaxAlarmes) THEN
    AlarmArray[AlarmCount] := '[M3] Defaut variateur translation AC600'; AlarmCount := AlarmCount + 1;
END_IF;
IF ((TranslationMotionErrorId AND 16#0040) <> 16#0000) AND (AlarmCount < CST_NbMaxAlarmes) THEN
    AlarmArray[AlarmCount] := '[M3] Limite extreme translation atteinte'; AlarmCount := AlarmCount + 1;
END_IF;
IF (TranslationFinalInterlockErrorId <> 16#0000) AND (AlarmCount < CST_NbMaxAlarmes) THEN
    AlarmArray[AlarmCount] := '[M3] Barriere finale translation (frein / redemarrage) - Reset'; AlarmCount := AlarmCount + 1;
END_IF;

// 5d. Collecte — benne (FB_Bucket.ErrorId, bits décodés)
//    Mapping = index cause FB_Bucket (FB_FaultCore : bit i = cause i) :
//    bit0 config géométrie · bit1 écart max · bit2 timeout · bit3 glissement M1 · bit4 codeurs non référencés
IF ((BucketErrorId AND 16#0001) <> 16#0000) AND (AlarmCount < CST_NbMaxAlarmes) THEN
    AlarmArray[AlarmCount] := '[BENNE] ErrorID:01 - configuration geometrie invalide'; AlarmCount := AlarmCount + 1;
END_IF;
IF ((BucketErrorId AND 16#0002) <> 16#0000) AND (AlarmCount < CST_NbMaxAlarmes) THEN
    AlarmArray[AlarmCount] := '[BENNE] ErrorID:02 - depassement ecart max autorise'; AlarmCount := AlarmCount + 1;
END_IF;
IF ((BucketErrorId AND 16#0004) <> 16#0000) AND EncM1Valid AND EncM2Valid AND (AlarmCount < CST_NbMaxAlarmes) THEN
    AlarmArray[AlarmCount] := '[BENNE] ErrorID:03 - timeout commande deplacement'; AlarmCount := AlarmCount + 1;
END_IF;
IF ((BucketErrorId AND 16#0008) <> 16#0000) AND (AlarmCount < CST_NbMaxAlarmes) THEN
    AlarmArray[AlarmCount] := '[BENNE] ErrorID:04 - glissement treuil M1'; AlarmCount := AlarmCount + 1;
END_IF;
IF ((BucketErrorId AND 16#0010) <> 16#0000) AND (AlarmCount < CST_NbMaxAlarmes) THEN
    AlarmArray[AlarmCount] := '[BENNE] ErrorID:05 - codeurs treuils non references'; AlarmCount := AlarmCount + 1;
END_IF;

// 5e. Collecte — synchro M1/M2 (FB_WinchSync.ErrorId)
IF ((SyncErrorId AND 16#0001) <> 16#0000) AND EncM1Valid AND EncM2Valid AND (AlarmCount < CST_NbMaxAlarmes) THEN
    AlarmArray[AlarmCount] := '[SYNC] ErrorID:01 - ecart M1/M2'; AlarmCount := AlarmCount + 1;
END_IF;
IF ((SyncErrorId AND 16#0002) <> 16#0000) AND (AlarmCount < CST_NbMaxAlarmes) THEN
    AlarmArray[AlarmCount] := '[SYNC] ErrorID:02 - incoherence commande'; AlarmCount := AlarmCount + 1;
END_IF;
// Discordance contacteurs M1/M2 decodee (FB_SyncContactor PRG_06 §2quinquies) : quel contacteur + niveau.
IF (SyncContactorDiag.MismatchLevel >= 1) AND (AlarmCount < CST_NbMaxAlarmes) THEN
    IF    SyncContactorDiag.RelayFwdMismatch THEN BannerSyncContactorWhich := 'relais montee';
    ELSIF SyncContactorDiag.RelayRevMismatch THEN BannerSyncContactorWhich := 'relais descente';
    ELSIF SyncContactorDiag.Step1Mismatch   THEN BannerSyncContactorWhich := 'palier 1';
    ELSIF SyncContactorDiag.Step2Mismatch   THEN BannerSyncContactorWhich := 'palier 2';
    ELSIF SyncContactorDiag.Step3Mismatch   THEN BannerSyncContactorWhich := 'palier 3';
    ELSIF SyncContactorDiag.Step4Mismatch   THEN BannerSyncContactorWhich := 'palier 4';
    ELSE  BannerSyncContactorWhich := 'non identifie';
    END_IF;
    IF SyncContactorDiag.MismatchLevel >= 2 THEN
        AlarmArray[AlarmCount] := CONCAT('[SYNC] discordance M1/M2 persistante -> coupure : ', BannerSyncContactorWhich);
    ELSE
        AlarmArray[AlarmCount] := CONCAT('[SYNC] discordance contacteurs M1/M2 -> arret : ', BannerSyncContactorWhich);
    END_IF;
    AlarmCount := AlarmCount + 1;
END_IF;

// 5f. Collecte — plongée / extraction (FB_DiveSearch / FB_ExtractionAssist)
IF ((DiveErrorId AND 16#0001) <> 16#0000) AND (AlarmCount < CST_NbMaxAlarmes) THEN
    AlarmArray[AlarmCount] := '[DIVE] ErrorID:01 - timeout immersion'; AlarmCount := AlarmCount + 1;
END_IF;
IF ((DiveErrorId AND 16#0002) <> 16#0000) AND (AlarmCount < CST_NbMaxAlarmes) THEN
    AlarmArray[AlarmCount] := '[DIVE] ErrorID:02 - timeout fond'; AlarmCount := AlarmCount + 1;
END_IF;
IF ((DiveErrorId AND 16#0004) <> 16#0000) AND EncM1Valid AND (AlarmCount < CST_NbMaxAlarmes) THEN
    AlarmArray[AlarmCount] := '[DIVE] ErrorID:03 - limite basse atteinte'; AlarmCount := AlarmCount + 1;
END_IF;
IF ((DiveErrorId AND 16#0008) <> 16#0000) AND (AlarmCount < CST_NbMaxAlarmes) THEN
    AlarmArray[AlarmCount] := '[DIVE] ErrorID:04 - contact fond perdu'; AlarmCount := AlarmCount + 1;
END_IF;
IF ((DiveErrorId AND 16#0010) <> 16#0000) AND (AlarmCount < CST_NbMaxAlarmes) THEN
    AlarmArray[AlarmCount] := '[DIVE] ErrorID:05 - perte tension cable'; AlarmCount := AlarmCount + 1;
END_IF;
IF ((DiveErrorId AND 16#0020) <> 16#0000) AND (AlarmCount < CST_NbMaxAlarmes) THEN
    AlarmArray[AlarmCount] := '[DIVE] ErrorID:06 - anomalie vitesse'; AlarmCount := AlarmCount + 1;
END_IF;
IF ((DiveErrorId AND 16#0040) <> 16#0000) AND (AlarmCount < CST_NbMaxAlarmes) THEN
    AlarmArray[AlarmCount] := '[DIVE] ErrorID:07 - config invalide'; AlarmCount := AlarmCount + 1;
END_IF;
IF ((ExtractionErrorId AND 16#0001) <> 16#0000) AND LocalIoValid AND (AlarmCount < CST_NbMaxAlarmes) THEN
    AlarmArray[AlarmCount] := '[EXTRACTION] ErrorID:01 - fond'; AlarmCount := AlarmCount + 1;
END_IF;
IF ((ExtractionErrorId AND 16#0002) <> 16#0000) AND (AlarmCount < CST_NbMaxAlarmes) THEN
    AlarmArray[AlarmCount] := '[EXTRACTION] ErrorID:02 - fermeture'; AlarmCount := AlarmCount + 1;
END_IF;
IF ((ExtractionErrorId AND 16#0004) <> 16#0000) AND (AlarmCount < CST_NbMaxAlarmes) THEN
    AlarmArray[AlarmCount] := '[EXTRACTION] ErrorID:03 - controle'; AlarmCount := AlarmCount + 1;
END_IF;
IF ((ExtractionErrorId AND 16#0008) <> 16#0000) AND (AlarmCount < CST_NbMaxAlarmes) THEN
    AlarmArray[AlarmCount] := '[EXTRACTION] ErrorID:04 - config'; AlarmCount := AlarmCount + 1;
END_IF;

// 5g. Collecte — AU / armement (FB_Safety_EmergencyManagement.Diag.ErrorId)
IF ((EmergencyErrorId AND 16#0001) <> 16#0000) AND (AlarmCount < CST_NbMaxAlarmes) THEN
    AlarmArray[AlarmCount] := '[AU] ErrorID:01 - redondance contacteurs'; AlarmCount := AlarmCount + 1;
END_IF;
IF ((EmergencyErrorId AND 16#0002) <> 16#0000) AND (AlarmCount < CST_NbMaxAlarmes) THEN
    AlarmArray[AlarmCount] := '[AU] ErrorID:02 - echec confirmation armement'; AlarmCount := AlarmCount + 1;
END_IF;
IF ((EmergencyErrorId AND 16#0008) <> 16#0000) AND (AlarmCount < CST_NbMaxAlarmes) THEN
    AlarmArray[AlarmCount] := '[AU] ErrorID:04 - echec autotest demarrage'; AlarmCount := AlarmCount + 1;
END_IF;

// 5h. Collecte — cycle semi-auto (FB_CycleSemiAuto.ErrorId)
IF ((CycleErrorId AND 16#0001) <> 16#0000) AND EncM1Valid AND (AlarmCount < CST_NbMaxAlarmes) THEN
    AlarmArray[AlarmCount] := '[CYCLE] ErrorID:01 - limite legale atteinte'; AlarmCount := AlarmCount + 1;
END_IF;
IF ((CycleErrorId AND 16#0002) <> 16#0000) AND EncM1Valid AND EncM2Valid AND (AlarmCount < CST_NbMaxAlarmes) THEN
    AlarmArray[AlarmCount] := '[CYCLE] ErrorID:02 - defaut synchro treuils'; AlarmCount := AlarmCount + 1;
END_IF;
IF ((CycleErrorId AND 16#0004) <> 16#0000) AND EncM1Valid AND EncM2Valid AND (AlarmCount < CST_NbMaxAlarmes) THEN
    AlarmArray[AlarmCount] := '[CYCLE] ErrorID:03 - ecart vitesse montee'; AlarmCount := AlarmCount + 1;
END_IF;
IF ((CycleErrorId AND 16#0008) <> 16#0000) AND (AlarmCount < CST_NbMaxAlarmes) THEN
    AlarmArray[AlarmCount] := '[CYCLE] ErrorID:04 - perte communication IHM'; AlarmCount := AlarmCount + 1;
END_IF;
IF ((CycleErrorId AND 16#0010) <> 16#0000) AND (AlarmCount < CST_NbMaxAlarmes) THEN
    AlarmArray[AlarmCount] := '[CYCLE] ErrorID:05 - timeout etape'; AlarmCount := AlarmCount + 1;
END_IF;
IF ((CycleErrorId AND 16#0020) <> 16#0000) AND EncM1Valid AND EncM2Valid AND (AlarmCount < CST_NbMaxAlarmes) THEN
    AlarmArray[AlarmCount] := '[CYCLE] ErrorID:06 - ecart codeurs remontee'; AlarmCount := AlarmCount + 1;
END_IF;
IF ((CycleErrorId AND 16#0080) <> 16#0000) AND (AlarmCount < CST_NbMaxAlarmes) THEN
    AlarmArray[AlarmCount] := '[CYCLE] ErrorID:08 - hors FDC haut translation P1'; AlarmCount := AlarmCount + 1;
END_IF;
IF ((CycleErrorId AND 16#0100) <> 16#0000) AND (AlarmCount < CST_NbMaxAlarmes) THEN
    AlarmArray[AlarmCount] := '[CYCLE] ErrorID:09 - palier 5 interdit en plongee'; AlarmCount := AlarmCount + 1;
END_IF;
IF ((CycleErrorId AND 16#0200) <> 16#0000) AND (AlarmCount < CST_NbMaxAlarmes) THEN
    AlarmArray[AlarmCount] := '[CYCLE] ErrorID:10 - palier 4 non confirme Kobold'; AlarmCount := AlarmCount + 1;
END_IF;
IF ((CycleErrorId AND 16#0800) <> 16#0000) AND (AlarmCount < CST_NbMaxAlarmes) THEN
    AlarmArray[AlarmCount] := '[CYCLE] ErrorID:12 - consigne profondeur invalide'; AlarmCount := AlarmCount + 1;
END_IF;

// 5h-bis. Collecte — defauts homing / commande treuils / codeurs / joystick / AU global
IF MachineHomingFailed AND (AlarmCount < CST_NbMaxAlarmes) THEN
    AlarmArray[AlarmCount] := '[HOMING] Echec ou abandon referencement machine - Reset'; AlarmCount := AlarmCount + 1;
END_IF;
IF MachineHomingLoss AND (AlarmCount < CST_NbMaxAlarmes) THEN
    AlarmArray[AlarmCount] := '[HOMING] Perte reference en mouvement - Reset'; AlarmCount := AlarmCount + 1;
END_IF;
IF WinchM1Error AND (AlarmCount < CST_NbMaxAlarmes) THEN
    AlarmArray[AlarmCount] := '[M1] Defaut commande ou barriere finale treuil'; AlarmCount := AlarmCount + 1;
END_IF;
IF WinchM2Error AND (AlarmCount < CST_NbMaxAlarmes) THEN
    AlarmArray[AlarmCount] := '[M2] Defaut commande ou barriere finale treuil'; AlarmCount := AlarmCount + 1;
END_IF;
IF EncoderM1Fault AND (AlarmCount < CST_NbMaxAlarmes) THEN
    AlarmArray[AlarmCount] := '[CODEUR] Defaut codeur treuil M1'; AlarmCount := AlarmCount + 1;
END_IF;
IF EncoderM2Fault AND (AlarmCount < CST_NbMaxAlarmes) THEN
    AlarmArray[AlarmCount] := '[CODEUR] Defaut codeur treuil M2'; AlarmCount := AlarmCount + 1;
END_IF;
IF JoystickLatchedFault AND (AlarmCount < CST_NbMaxAlarmes) THEN
    AlarmArray[AlarmCount] := '[JOYSTICK] Defaut joystick latche - Reset'; AlarmCount := AlarmCount + 1;
END_IF;
IF SyncFaultLatched AND ((SyncErrorId AND 16#0003) = 16#0000) AND (AlarmCount < CST_NbMaxAlarmes) THEN
    AlarmArray[AlarmCount] := '[SYNC] Defaut synchro treuils latche - Reset'; AlarmCount := AlarmCount + 1;
END_IF;
IF BucketFaultLatched AND ((BucketErrorId AND 16#001F) = 16#0000) AND (AlarmCount < CST_NbMaxAlarmes) THEN
    AlarmArray[AlarmCount] := '[BENNE] Defaut benne latche - Reset'; AlarmCount := AlarmCount + 1;
END_IF;
